screen "8_1" 800x480, template "Template_2"
   Button "Button_1" at 40,240 size 120x40; TextOff 'Acyclovir'
      on Click: ActivateScreen("4_ORDER", 0); SetTag("Selected_URL", 'file:///C:/ASRS_Video/clip291.html')
      on Activate: SetTag("Selected_Medicine", 291)
      on Release: SetTag("ยา 291", 0)
      on Press: SetTag("ยา 291", 1)
   Button "Button_10" at 40,416 size 120x40; TextOff 'Remdesivir'
      on Click: ActivateScreen("4_ORDER", 0); SetTag("Selected_URL", 'file:///C:/ASRS_Video/clip296.html')
      on Activate: SetTag("Selected_Medicine", 296)
      on Release: SetTag("ยา 296", 0)
      on Press: SetTag("ยา 296", 1)
   Button "Button_2" at 191,241 size 120x40; TextOff 'Valacyclovir'
      on Click: ActivateScreen("4_ORDER", 0); SetTag("Selected_URL", 'file:///C:/ASRS_Video/clip292.html')
      on Activate: SetTag("Selected_Medicine", 292)
      on Release: SetTag("ยา 292", 0)
      on Press: SetTag("ยา 292", 1)
   Button "Button_3" at 192,416 size 120x40; TextOff 'Favipiravir'
      on Click: ActivateScreen("4_ORDER", 0); SetTag("Selected_URL", 'file:///C:/ASRS_Video/clip297.html')
      on Activate: SetTag("Selected_Medicine", 297)
      on Release: SetTag("ยา 297", 0)
      on Press: SetTag("ยา 297", 1)
   Button "Button_4" at 342,241 size 120x40; TextOff 'Ganciclovir'
      on Click: ActivateScreen("4_ORDER", 0); SetTag("Selected_URL", 'file:///C:/ASRS_Video/clip293.html')
      on Activate: SetTag("Selected_Medicine", 293)
      on Release: SetTag("ยา 293", 0)
      on Press: SetTag("ยา 293", 1)
   Button "Button_5" at 342,417 size 120x40; TextOff 'Lamivudine'
      on Click: ActivateScreen("4_ORDER", 0); SetTag("Selected_URL", 'file:///C:/ASRS_Video/clip298.html')
      on Activate: SetTag("Selected_Medicine", 298)
      on Release: SetTag("ยา 298", 0)
      on Press: SetTag("ยา 298", 1)
   Button "Button_6" at 492,416 size 120x40; TextOff 'Zidovudine'
      on Click: ActivateScreen("4_ORDER", 0); SetTag("Selected_URL", 'file:///C:/ASRS_Video/clip299.html')
      on Activate: SetTag("Selected_Medicine", 299)
      on Release: SetTag("ยา 299", 0)
      on Press: SetTag("ยา 299", 1)
   Button "Button_7" at 492,240 size 120x40; TextOff 'Oseltamivir'
      on Click: ActivateScreen("4_ORDER", 0); SetTag("Selected_URL", 'file:///C:/ASRS_Video/clip294.html')
      on Activate: SetTag("Selected_Medicine", 294)
      on Release: SetTag("ยา 294", 0)
      on Press: SetTag("ยา 294", 1)
   Button "Button_8" at 644,240 size 120x40; TextOff 'Zanamivir'
      on Click: ActivateScreen("4_ORDER", 0); SetTag("Selected_URL", 'file:///C:/ASRS_Video/clip295.html')
      on Activate: SetTag("Selected_Medicine", 295)
      on Release: SetTag("ยา 295", 0)
      on Press: SetTag("ยา 295", 1)
   Button "Button_11" at 645,416 size 120x40; TextOff 'Tenofovir'
      on Click: ActivateScreen("4_ORDER", 0); SetTag("Selected_URL", 'file:///C:/ASRS_Video/clip300.html')
      on Activate: SetTag("Selected_Medicine", 300)
      on Release: SetTag("ยา 300", 0)
      on Press: SetTag("ยา 300", 1)
   Button "Button_12" at 24,16 size 94x40; TextOff 'Back'
      on Press: ActivateScreen("7_1", 0)
   Button "Button_9" at 688,16 size 96x40; TextOff 'Next'
      on Press: ActivateScreen("9_1", 0)
   GraphicView "Template_Graphic view_2" at 27,19 size 36x32; Picture "fast-backward"
   GraphicView "Template_Graphic view_1" at 693,20 size 36x32; Picture "play"
   GraphicView "Template_Graphic view_3" at 37,128 size 120x104; Picture "71"
   GraphicView "Template_Graphic view_4" at 191,129 size 120x104; Picture "72"
   GraphicView "Template_Graphic view_5" at 339,129 size 120x104; Picture "73"
   GraphicView "Template_Graphic view_6" at 493,129 size 120x104; Picture "74"
   GraphicView "Template_Graphic view_7" at 645,129 size 120x104; Picture "75"
   GraphicView "Template_Graphic view_8" at 38,305 size 120x104; Picture "76"
   GraphicView "Template_Graphic view_9" at 189,304 size 120x112; Picture "77"
   GraphicView "Template_Graphic view_10" at 351,307 size 96x104; Picture "78"
   GraphicView "Template_Graphic view_11" at 491,299 size 120x112; Picture "79"
   GraphicView "Template_Graphic view_12" at 645,304 size 120x104; Picture "80"
   TextField "Template_Text field_2" at 201,80 size 20x32; Text '8'

screen "9_1" 800x480, template "Template_2"
   Button "Button_1" at 38,239 size 120x40; TextOff 'Efavirenz'
      on Click: ActivateScreen("4_ORDER", 0); SetTag("Selected_URL", 'file:///C:/ASRS_Video/clip301.html')
      on Activate: SetTag("Selected_Medicine", 301)
      on Release: SetTag("ยา 301", 0)
      on Press: SetTag("ยา 301", 1)
   Button "Button_10" at 38,415 size 120x40; TextOff 'Mebendazole'
      on Click: ActivateScreen("4_ORDER", 0); SetTag("Selected_URL", 'file:///C:/ASRS_Video/clip306.html')
      on Activate: SetTag("Selected_Medicine", 306)
      on Release: SetTag("ยา 306", 0)
      on Press: SetTag("ยา 306", 1)
   Button "Button_2" at 189,240 size 120x40; TextOff 'Dolutegravir'
      on Click: ActivateScreen("4_ORDER", 0); SetTag("Selected_URL", 'file:///C:/ASRS_Video/clip302.html')
      on Activate: SetTag("Selected_Medicine", 302)
      on Release: SetTag("ยา 302", 0)
      on Press: SetTag("ยา 302", 1)
   Button "Button_3" at 190,415 size 120x40; TextOff 'Ivermectin'
      on Click: ActivateScreen("4_ORDER", 0); SetTag("Selected_URL", 'file:///C:/ASRS_Video/clip307.html')
      on Activate: SetTag("Selected_Medicine", 307)
      on Release: SetTag("ยา 307", 0)
      on Press: SetTag("ยา 307", 1)
   Button "Button_4" at 340,240 size 120x40; TextOff 'Nevirapine'
      on Click: ActivateScreen("4_ORDER", 0); SetTag("Selected_URL", 'file:///C:/ASRS_Video/clip303.html')
      on Activate: SetTag("Selected_Medicine", 303)
      on Release: SetTag("ยา 303", 0)
      on Press: SetTag("ยา 303", 1)
   Button "Button_5" at 340,416 size 120x40; TextOff 'Praziquantel'
      on Click: ActivateScreen("4_ORDER", 0); SetTag("Selected_URL", 'file:///C:/ASRS_Video/clip308.html')
      on Activate: SetTag("Selected_Medicine", 308)
      on Release: SetTag("ยา 308", 0)
      on Press: SetTag("ยา 308", 1)
   Button "Button_6" at 492,416 size 120x40; TextOff 'Pyrantel pamoate'
      on Click: ActivateScreen("4_ORDER", 0); SetTag("Selected_URL", 'file:///C:/ASRS_Video/clip309.html')
      on Activate: SetTag("Selected_Medicine", 309)
      on Release: SetTag("ยา 309", 0)
      on Press: SetTag("ยา 309", 1)
   Button "Button_7" at 492,240 size 120x40; TextOff 'Lopinavir ritonavir'
      on Click: ActivateScreen("4_ORDER", 0); SetTag("Selected_URL", 'file:///C:/ASRS_Video/clip304.html')
      on Activate: SetTag("Selected_Medicine", 304)
      on Release: SetTag("ยา 304", 0)
      on Press: SetTag("ยา 304", 1)
   Button "Button_8" at 644,240 size 120x40; TextOff 'Albendazole'
      on Click: ActivateScreen("4_ORDER", 0); SetTag("Selected_URL", 'file:///C:/ASRS_Video/clip305.html')
      on Activate: SetTag("Selected_Medicine", 305)
      on Release: SetTag("ยา 305", 0)
      on Press: SetTag("ยา 305", 1)
   Button "Button_11" at 645,416 size 120x40; TextOff 'Diethylcarbamazine'
      on Click: ActivateScreen("4_ORDER", 0); SetTag("Selected_URL", 'file:///C:/ASRS_Video/clip310.html')
      on Activate: SetTag("Selected_Medicine", 310)
      on Release: SetTag("ยา 310", 0)
      on Press: SetTag("ยา 310", 1)
   Button "Button_12" at 24,16 size 94x40; TextOff 'Back'
      on Press: ActivateScreen("8_1", 0)
   Button "Button_9" at 688,16 size 96x40; TextOff 'Next'
      on Press: ActivateScreen("10_1", 0)
   GraphicView "Template_Graphic view_2" at 27,19 size 36x32; Picture "fast-backward"
   GraphicView "Template_Graphic view_1" at 693,20 size 36x32; Picture "play"
   GraphicView "Template_Graphic view_3" at 37,128 size 120x104; Picture "81"
   GraphicView "Template_Graphic view_4" at 191,129 size 120x104; Picture "82"
   GraphicView "Template_Graphic view_5" at 339,129 size 120x104; Picture "83"
   GraphicView "Template_Graphic view_6" at 493,129 size 120x104; Picture "84"
   GraphicView "Template_Graphic view_7" at 645,129 size 120x104; Picture "85"
   GraphicView "Template_Graphic view_8" at 38,305 size 120x104; Picture "86"
   GraphicView "Template_Graphic view_9" at 189,304 size 120x112; Picture "87"
   GraphicView "Template_Graphic view_10" at 351,307 size 96x104; Picture "88"
   GraphicView "Template_Graphic view_11" at 497,304 size 120x112; Picture "89"
   GraphicView "Template_Graphic view_12" at 645,304 size 120x104; Picture "90"
   TextField "Template_Text field_2" at 201,80 size 20x32; Text '9'

screen "10_1" 800x480, template "Template_2"
   Button "Button_1" at 38,239 size 120x40; TextOff 'Chloroquine'
      on Click: ActivateScreen("4_ORDER", 0); SetTag("Selected_URL", 'file:///C:/ASRS_Video/clip311.html')
      on Activate: SetTag("Selected_Medicine", 311)
      on Release: SetTag("ยา 311", 0)
      on Press: SetTag("ยา 311", 1)
   Button "Button_10" at 38,415 size 120x40; TextOff 'Dapsone'
      on Click: ActivateScreen("4_ORDER", 0); SetTag("Selected_URL", 'file:///C:/ASRS_Video/clip316.html')
      on Activate: SetTag("Selected_Medicine", 316)
      on Release: SetTag("ยา 316", 0)
      on Press: SetTag("ยา 316", 1)
   Button "Button_2" at 189,240 size 120x40; TextOff 'Primaquine'
      on Click: ActivateScreen("4_ORDER", 0); SetTag("Selected_URL", 'file:///C:/ASRS_Video/clip312.html')
      on Activate: SetTag("Selected_Medicine", 312)
      on Release: SetTag("ยา 312", 0)
      on Press: SetTag("ยา 312", 1)
   Button "Button_3" at 190,415 size 120x40; TextOff 'Permethrin'
      on Click: ActivateScreen("4_ORDER", 0); SetTag("Selected_URL", 'file:///C:/ASRS_Video/clip317.html')
      on Activate: SetTag("Selected_Medicine", 317)
      on Release: SetTag("ยา 317", 0)
      on Press: SetTag("ยา 317", 1)
   Button "Button_4" at 340,240 size 120x40; TextOff 'Artesunate'
      on Click: ActivateScreen("4_ORDER", 0); SetTag("Selected_URL", 'file:///C:/ASRS_Video/clip313.html')
      on Activate: SetTag("Selected_Medicine", 313)
      on Release: SetTag("ยา 313", 0)
      on Press: SetTag("ยา 313", 1)
   Button "Button_5" at 340,416 size 120x40; TextOff 'Benzyl benzoate'
      on Click: ActivateScreen("4_ORDER", 0); SetTag("Selected_URL", 'file:///C:/ASRS_Video/clip318.html')
      on Activate: SetTag("Selected_Medicine", 318)
      on Release: SetTag("ยา 318", 0)
      on Press: SetTag("ยา 318", 1)
   Button "Button_6" at 492,416 size 120x40; TextOff 'Povidone iodine'
      on Click: ActivateScreen("4_ORDER", 0); SetTag("Selected_URL", 'file:///C:/ASRS_Video/clip319.html')
      on Activate: SetTag("Selected_Medicine", 319)
      on Release: SetTag("ยา 319", 0)
      on Press: SetTag("ยา 319", 1)
   Button "Button_7" at 492,240 size 120x40; TextOff 'Artemether lumefantrine'
      on Click: ActivateScreen("4_ORDER", 0); SetTag("Selected_URL", 'file:///C:/ASRS_Video/clip314.html')
      on Activate: SetTag("Selected_Medicine", 314)
      on Release: SetTag("ยา 314", 0)
      on Press: SetTag("ยา 314", 1)
   Button "Button_8" at 644,240 size 120x40; TextOff 'Quinine'
      on Click: ActivateScreen("4_ORDER", 0); SetTag("Selected_URL", 'file:///C:/ASRS_Video/clip315.html')
      on Activate: SetTag("Selected_Medicine", 315)
      on Release: SetTag("ยา 315", 0)
      on Press: SetTag("ยา 315", 1)
   Button "Button_11" at 645,416 size 120x40; TextOff 'Chlorhexidine'
      on Click: ActivateScreen("4_ORDER", 0); SetTag("Selected_URL", 'file:///C:/ASRS_Video/clip320.html')
      on Activate: SetTag("Selected_Medicine", 320)
      on Release: SetTag("ยา 320", 0)
      on Press: SetTag("ยา 320", 1)
   Button "Button_12" at 24,16 size 94x40; TextOff 'Back'
      on Press: ActivateScreen("9_1", 0)
   Button "Button_9" at 688,16 size 96x40; TextOff 'Next'
      on Press: ActivateScreen("11_1", 0)
   GraphicView "Template_Graphic view_2" at 27,19 size 36x32; Picture "fast-backward"
   GraphicView "Template_Graphic view_1" at 693,20 size 36x32; Picture "play"
   GraphicView "Template_Graphic view_3" at 37,128 size 120x104; Picture "91"
   GraphicView "Template_Graphic view_4" at 191,129 size 120x104; Picture "92"
   GraphicView "Template_Graphic view_5" at 339,129 size 120x104; Picture "93"
   GraphicView "Template_Graphic view_6" at 493,129 size 120x104; Picture "94"
   GraphicView "Template_Graphic view_7" at 645,129 size 120x104; Picture "95"
   GraphicView "Template_Graphic view_8" at 38,305 size 120x104; Picture "96"
   GraphicView "Template_Graphic view_9" at 189,304 size 120x112; Picture "97"
   GraphicView "Template_Graphic view_10" at 351,307 size 96x104; Picture "98"
   GraphicView "Template_Graphic view_11" at 497,304 size 104x104; Picture "99"
   GraphicView "Template_Graphic view_12" at 645,304 size 120x104; Picture "100"
   TextField "Template_Text field_2" at 201,80 size 36x32; Text '10'

screen "11_1" 800x480, template "Template_2"
   Button "Button_1" at 38,239 size 120x40; TextOff 'Colistin'
      on Click: ActivateScreen("4_ORDER", 0); SetTag("Selected_URL", 'file:///C:/ASRS_Video/clip321.html')
      on Activate: SetTag("Selected_Medicine", 321)
      on Release: SetTag("ยา 321", 0)
      on Press: SetTag("ยา 321", 1)
   Button "Button_10" at 38,415 size 120x40; TextOff 'Rabies vaccine'
      on Click: ActivateScreen("4_ORDER", 0); SetTag("Selected_URL", 'file:///C:/ASRS_Video/clip326.html')
      on Activate: SetTag("Selected_Medicine", 326)
      on Release: SetTag("ยา 326", 0)
      on Press: SetTag("ยา 326", 1)
   Button "Button_2" at 189,240 size 120x40; TextOff 'Caspofungin'
      on Click: ActivateScreen("4_ORDER", 0); SetTag("Selected_URL", 'file:///C:/ASRS_Video/clip322.html')
      on Activate: SetTag("Selected_Medicine", 322)
      on Release: SetTag("ยา 322", 0)
      on Press: SetTag("ยา 322", 1)
   Button "Button_3" at 190,415 size 120x40; TextOff 'Influenza vaccine'
      on Click: ActivateScreen("4_ORDER", 0); SetTag("Selected_URL", 'file:///C:/ASRS_Video/clip327.html')
      on Activate: SetTag("Selected_Medicine", 327)
      on Release: SetTag("ยา 327", 0)
      on Press: SetTag("ยา 327", 1)
   Button "Button_4" at 340,240 size 120x40; TextOff 'Bacitracin'
      on Click: ActivateScreen("4_ORDER", 0); SetTag("Selected_URL", 'file:///C:/ASRS_Video/clip323.html')
      on Activate: SetTag("Selected_Medicine", 323)
      on Release: SetTag("ยา 323", 0)
      on Press: SetTag("ยา 323", 1)
   Button "Button_5" at 340,416 size 120x40; TextOff 'Hepatitis B vaccine'
      on Click: ActivateScreen("4_ORDER", 0); SetTag("Selected_URL", 'file:///C:/ASRS_Video/clip328.html')
      on Activate: SetTag("Selected_Medicine", 328)
      on Release: SetTag("ยา 328", 0)
      on Press: SetTag("ยา 328", 1)
   Button "Button_6" at 492,416 size 120x40; TextOff 'BCG vaccine'
      on Click: ActivateScreen("4_ORDER", 0); SetTag("Selected_URL", 'file:///C:/ASRS_Video/clip329.html')
      on Activate: SetTag("Selected_Medicine", 329)
      on Release: SetTag("ยา 329", 0)
      on Press: SetTag("ยา 329", 1)
   Button "Button_7" at 492,240 size 120x40; TextOff 'Fusidic acid'
      on Click: ActivateScreen("4_ORDER", 0); SetTag("Selected_URL", 'file:///C:/ASRS_Video/clip324.html')
      on Activate: SetTag("Selected_Medicine", 324)
      on Release: SetTag("ยา 324", 0)
      on Press: SetTag("ยา 324", 1)
   Button "Button_8" at 644,240 size 120x40; TextOff 'Mupirocin'
      on Click: ActivateScreen("4_ORDER", 0); SetTag("Selected_URL", 'file:///C:/ASRS_Video/clip325.html')
      on Activate: SetTag("Selected_Medicine", 325)
      on Release: SetTag("ยา 325", 0)
      on Press: SetTag("ยา 325", 1)
   Button "Button_11" at 645,416 size 120x40; TextOff 'DTP vaccine'
      on Click: ActivateScreen("4_ORDER", 0); SetTag("Selected_URL", 'file:///C:/ASRS_Video/clip330.html')
      on Activate: SetTag("Selected_Medicine", 330)
      on Release: SetTag("ยา 330", 0)
      on Press: SetTag("ยา 330", 1)
   Button "Button_12" at 24,16 size 94x40; TextOff 'Back'
      on Press: ActivateScreen("10_1", 0)
   Button "Button_9" at 688,16 size 96x40; TextOff 'Next'
      on Press: ActivateScreen("12_1", 0)
   GraphicView "Template_Graphic view_2" at 27,19 size 36x32; Picture "fast-backward"
   GraphicView "Template_Graphic view_1" at 693,20 size 36x32; Picture "play"
   GraphicView "Template_Graphic view_3" at 37,128 size 120x104; Picture "101"
   GraphicView "Template_Graphic view_4" at 191,129 size 120x104; Picture "102"
   GraphicView "Template_Graphic view_5" at 339,129 size 120x104; Picture "103"
   GraphicView "Template_Graphic view_6" at 493,129 size 120x104; Picture "104"
   GraphicView "Template_Graphic view_7" at 645,129 size 120x104; Picture "105"
   GraphicView "Template_Graphic view_8" at 38,305 size 120x104; Picture "106"
   GraphicView "Template_Graphic view_9" at 189,304 size 120x104; Picture "107"
   GraphicView "Template_Graphic view_10" at 351,307 size 96x104; Picture "108"
   GraphicView "Template_Graphic view_11" at 497,304 size 112x104; Picture "109"
   GraphicView "Template_Graphic view_12" at 645,304 size 120x104; Picture "110"
   TextField "Template_Text field_2" at 201,80 size 36x32; Text '11'

screen "12_1" 800x480, template "Template_2"
   Button "Button_1" at 38,239 size 120x40; TextOff 'MMR vaccine'
      on Click: ActivateScreen("4_ORDER", 0); SetTag("Selected_URL", 'file:///C:/ASRS_Video/clip331.html')
      on Activate: SetTag("Selected_Medicine", 331)
      on Release: SetTag("ยา 331", 0)
      on Press: SetTag("ยา 331", 1)
   Button "Button_10" at 38,415 size 120x40; TextOff 'Rotavirus vaccine'
      on Click: ActivateScreen("4_ORDER", 0); SetTag("Selected_URL", 'file:///C:/ASRS_Video/clip336.html')
      on Activate: SetTag("Selected_Medicine", 336)
      on Release: SetTag("ยา 336", 0)
      on Press: SetTag("ยา 336", 1)
   Button "Button_2" at 189,240 size 120x40; TextOff 'JE vaccine'
      on Click: ActivateScreen("4_ORDER", 0); SetTag("Selected_URL", 'file:///C:/ASRS_Video/clip332.html')
      on Activate: SetTag("Selected_Medicine", 332)
      on Release: SetTag("ยา 332", 0)
      on Press: SetTag("ยา 332", 1)
   Button "Button_3" at 190,415 size 120x40; TextOff 'COVID-19 vaccine'
      on Click: ActivateScreen("4_ORDER", 0); SetTag("Selected_URL", 'file:///C:/ASRS_Video/clip337.html')
      on Activate: SetTag("Selected_Medicine", 337)
      on Release: SetTag("ยา 337", 0)
      on Press: SetTag("ยา 337", 1)
   Button "Button_4" at 340,240 size 120x40; TextOff 'HPV vaccine'
      on Click: ActivateScreen("4_ORDER", 0); SetTag("Selected_URL", 'file:///C:/ASRS_Video/clip333.html')
      on Activate: SetTag("Selected_Medicine", 333)
      on Release: SetTag("ยา 333", 0)
      on Press: SetTag("ยา 333", 1)
   Button "Button_5" at 340,416 size 120x40; TextOff 'Tetanus toxoid'
      on Click: ActivateScreen("4_ORDER", 0); SetTag("Selected_URL", 'file:///C:/ASRS_Video/clip338.html')
      on Activate: SetTag("Selected_Medicine", 338)
      on Release: SetTag("ยา 338", 0)
      on Press: SetTag("ยา 338", 1)
   Button "Button_6" at 492,416 size 120x40; TextOff 'Rabies immunoglobulin'
      on Click: ActivateScreen("4_ORDER", 0); SetTag("Selected_URL", 'file:///C:/ASRS_Video/clip339.html')
      on Activate: SetTag("Selected_Medicine", 339)
      on Release: SetTag("ยา 339", 0)
      on Press: SetTag("ยา 339", 1)
   Button "Button_7" at 492,240 size 120x40; TextOff 'Varicella vaccine'
      on Click: ActivateScreen("4_ORDER", 0); SetTag("Selected_URL", 'file:///C:/ASRS_Video/clip334.html')
      on Activate: SetTag("Selected_Medicine", 334)
      on Release: SetTag("ยา 334", 0)
      on Press: SetTag("ยา 334", 1)
   Button "Button_8" at 644,240 size 120x40; TextOff 'Pneumococcal vaccine'
      on Click: ActivateScreen("4_ORDER", 0); SetTag("Selected_URL", 'file:///C:/ASRS_Video/clip335.html')
      on Activate: SetTag("Selected_Medicine", 335)
      on Release: SetTag("ยา 335", 0)
      on Press: SetTag("ยา 335", 1)
   Button "Button_11" at 645,416 size 120x40; TextOff 'Hepatitis B immunoglobulin'
      on Click: ActivateScreen("4_ORDER", 0); SetTag("Selected_URL", 'file:///C:/ASRS_Video/clip340.html')
      on Activate: SetTag("Selected_Medicine", 340)
      on Release: SetTag("ยา 340", 0)
      on Press: SetTag("ยา 340", 1)
   Button "Button_12" at 24,16 size 94x40; TextOff 'Back'
      on Press: ActivateScreen("11_1", 0)
   GraphicView "Template_Graphic view_2" at 27,19 size 36x32; Picture "fast-backward"
   GraphicView "Template_Graphic view_3" at 37,128 size 120x104; Picture "111"
   GraphicView "Template_Graphic view_4" at 191,129 size 120x104; Picture "112"
   GraphicView "Template_Graphic view_5" at 339,129 size 120x104; Picture "113"
   GraphicView "Template_Graphic view_6" at 493,129 size 120x104; Picture "114"
   GraphicView "Template_Graphic view_7" at 645,129 size 120x104; Picture "115"
   GraphicView "Template_Graphic view_8" at 38,305 size 120x104; Picture "116"
   GraphicView "Template_Graphic view_9" at 189,304 size 120x112; Picture "117"
   GraphicView "Template_Graphic view_10" at 351,307 size 96x104; Picture "118"
   GraphicView "Template_Graphic view_11" at 497,304 size 120x112; Picture "119"
   GraphicView "Template_Graphic view_12" at 645,304 size 120x104; Picture "120"
   TextField "Template_Text field_2" at 201,80 size 36x32; Text '12'

screen "1-10" 800x480, template "Template_2"
   Button "Button_1" at 40,240 size 120x40; TextOff 'Lidocaine'
      on Click: ActivateScreen("4_ORDER", 0); SetTag("Selected_URL", 'file:///C:/ASRS_Video/clip1.html')
      on Activate: SetTag("Selected_Medicine", 1)
      on Release: SetTag("ยา 1", 0)
      on Press: SetTag("ยา 1", 1)
   Button "Button_10" at 38,415 size 120x40; TextOff 'Tetracaine'
      on Click: ActivateScreen("4_ORDER", 0); SetTag("Selected_URL", 'file:///C:/ASRS_Video/clip6.html')
      on Activate: SetTag("Selected_Medicine", 6)
      on Release: SetTag("ยา 6", 0)
      on Press: SetTag("ยา 6", 1)
   Button "Button_2" at 189,240 size 120x40; TextOff 'Bupivacaine'
      on Click: ActivateScreen("4_ORDER", 0); SetTag("Selected_URL", 'file:///C:/ASRS_Video/clip2.html')
      on Activate: SetTag("Selected_Medicine", 2)
      on Release: SetTag("ยา 2", 0)
      on Press: SetTag("ยา 2", 1)
   Button "Button_3" at 190,415 size 120x40; TextOff 'Propofol'
      on Click: ActivateScreen("4_ORDER", 0); SetTag("Selected_URL", 'file:///C:/ASRS_Video/clip7.html')
      on Activate: SetTag("Selected_Medicine", 7)
      on Release: SetTag("ยา 7", 0)
      on Press: SetTag("ยา 7", 1)
   Button "Button_4" at 340,240 size 120x40; TextOff 'Ropivacaine'
      on Click: ActivateScreen("4_ORDER", 0); SetTag("Selected_URL", 'file:///C:/ASRS_Video/clip3.html')
      on Activate: SetTag("Selected_Medicine", 3)
      on Release: SetTag("ยา 3", 0)
      on Press: SetTag("ยา 3", 1)
   Button "Button_5" at 340,416 size 120x40; TextOff 'Ketamine'
      on Click: ActivateScreen("4_ORDER", 0); SetTag("Selected_URL", 'file:///C:/ASRS_Video/clip8.html')
      on Activate: SetTag("Selected_Medicine", 8)
      on Release: SetTag("ยา 8", 0)
      on Press: SetTag("ยา 8", 1)
   Button "Button_6" at 492,416 size 120x40; TextOff 'Etomidate'
      on Click: ActivateScreen("4_ORDER", 0); SetTag("Selected_URL", 'file:///C:/ASRS_Video/clip9.html')
      on Activate: SetTag("Selected_Medicine", 9)
      on Release: SetTag("ยา 9", 0)
      on Press: SetTag("ยา 9", 1)
   Button "Button_7" at 492,240 size 120x40; TextOff 'Procaine'
      on Click: ActivateScreen("4_ORDER", 0); SetTag("Selected_URL", 'file:///C:/ASRS_Video/clip4.html')
      on Activate: SetTag("Selected_Medicine", 4)
      on Release: SetTag("ยา 4", 0)
      on Press: SetTag("ยา 4", 1)
   Button "Button_8" at 644,240 size 120x40; TextOff 'Benzocaine'
      on Click: ActivateScreen("4_ORDER", 0); SetTag("Selected_URL", 'file:///C:/ASRS_Video/clip5.html')
      on Activate: SetTag("Selected_Medicine", 5)
      on Release: SetTag("ยา 5", 0)
      on Press: SetTag("ยา 5", 1)
   Button "Button_11" at 645,416 size 120x40; TextOff 'Thiopental'
      on Click: ActivateScreen("4_ORDER", 0); SetTag("Selected_URL", 'file:///C:/ASRS_Video/clip10.html')
      on Activate: SetTag("Selected_Medicine", 10)
      on Release: SetTag("ยา 10", 0)
      on Press: SetTag("ยา 10", 1)
   Button "Button_12" at 688,16 size 96x40; TextOff 'Next'
      on Press: ActivateScreen("11-20", 0)
   Button "Button_9" at 24,16 size 94x40; TextOff 'Back'
      on Press: ActivateScreen("4_ORDER", 0)
   GraphicView "Template_Graphic view_2" at 693,20 size 36x32; Picture "play"
   GraphicView "Template_Graphic view_1" at 27,19 size 36x32; Picture "fast-backward"
   GraphicView "Template_Graphic view_3" at 38,127 size 120x112; Picture "Picture1"
   GraphicView "Template_Graphic view_4" at 190,128 size 120x112; Picture "Picture2"
   GraphicView "Template_Graphic view_5" at 340,128 size 120x112; Picture "Picture3"
   GraphicView "Template_Graphic view_6" at 493,128 size 120x112; Picture "Picture4"
   GraphicView "Template_Graphic view_7" at 644,128 size 120x112; Picture "Picture5"
   GraphicView "Template_Graphic view_8" at 37,302 size 120x112; Picture "Picture6"
   GraphicView "Template_Graphic view_9" at 189,303 size 120x112; Picture "Picture7"
   GraphicView "Template_Graphic view_10" at 339,303 size 120x112; Picture "Picture8"
   GraphicView "Template_Graphic view_11" at 492,303 size 120x112; Picture "Picture9"
   GraphicView "Template_Graphic view_12" at 643,303 size 120x112; Picture "Picture10"
   TextField "Template_Text field_2" at 201,80 size 20x32; Text '1'

screen "11-20" 800x480, template "Template_2"
   Button "Button_1" at 38,239 size 120x40; TextOff 'Midazolam'
      on Click: ActivateScreen("4_ORDER", 0); SetTag("Selected_URL", 'file:///C:/ASRS_Video/clip11.html')
      on Activate: SetTag("Selected_Medicine", 11)
      on Release: SetTag("ยา 11", 0)
      on Press: SetTag("ยา 11", 1)
   Button "Button_9" at 688,16 size 96x40; TextOff 'Next'
      on Press: ActivateScreen("21-30", 0)
   Button "Button_10" at 38,415 size 120x40; TextOff 'Pethidine'
      on Click: ActivateScreen("4_ORDER", 0); SetTag("Selected_URL", 'file:///C:/ASRS_Video/clip16.html')
      on Activate: SetTag("Selected_Medicine", 16)
      on Release: SetTag("ยา 16", 0)
      on Press: SetTag("ยา 16", 1)
   Button "Button_2" at 189,240 size 120x40; TextOff 'Diazepam'
      on Click: ActivateScreen("4_ORDER", 0); SetTag("Selected_URL", 'file:///C:/ASRS_Video/clip12.html')
      on Activate: SetTag("Selected_Medicine", 12)
      on Release: SetTag("ยา 12", 0)
      on Press: SetTag("ยา 12", 1)
   Button "Button_3" at 190,415 size 120x40; TextOff 'Tramadol'
      on Click: ActivateScreen("4_ORDER", 0); SetTag("Selected_URL", 'file:///C:/ASRS_Video/clip17.html')
      on Activate: SetTag("Selected_Medicine", 17)
      on Release: SetTag("ยา 17", 0)
      on Press: SetTag("ยา 17", 1)
   Button "Button_4" at 340,240 size 120x40; TextOff 'Lorazepam'
      on Click: ActivateScreen("4_ORDER", 0); SetTag("Selected_URL", 'file:///C:/ASRS_Video/clip13.html')
      on Activate: SetTag("Selected_Medicine", 13)
      on Release: SetTag("ยา 13", 0)
      on Press: SetTag("ยา 13", 1)
   Button "Button_5" at 340,416 size 120x40; TextOff 'Nalbuphine'
      on Click: ActivateScreen("4_ORDER", 0); SetTag("Selected_URL", 'file:///C:/ASRS_Video/clip18.html')
      on Activate: SetTag("Selected_Medicine", 18)
      on Release: SetTag("ยา 18", 0)
      on Press: SetTag("ยา 18", 1)
   Button "Button_6" at 492,416 size 120x40; TextOff 'Remifentanil'
      on Click: ActivateScreen("4_ORDER", 0); SetTag("Selected_URL", 'file:///C:/ASRS_Video/clip19.html')
      on Activate: SetTag("Selected_Medicine", 19)
      on Release: SetTag("ยา 19", 0)
      on Press: SetTag("ยา 19", 1)
   Button "Button_7" at 492,240 size 120x40; TextOff 'Fentanyl'
      on Click: ActivateScreen("4_ORDER", 0); SetTag("Selected_URL", 'file:///C:/ASRS_Video/clip14.html')
      on Activate: SetTag("Selected_Medicine", 14)
      on Release: SetTag("ยา 14", 0)
      on Press: SetTag("ยา 14", 1)
   Button "Button_8" at 644,240 size 120x40; TextOff 'Morphine'
      on Click: ActivateScreen("4_ORDER", 0); SetTag("Selected_URL", 'file:///C:/ASRS_Video/clip15.html')
      on Activate: SetTag("Selected_Medicine", 15)
      on Release: SetTag("ยา 15", 0)
      on Press: SetTag("ยา 15", 1)
   Button "Button_11" at 645,416 size 120x40; TextOff 'Succinylcholine'
      on Click: ActivateScreen("4_ORDER", 0); SetTag("Selected_URL", 'file:///C:/ASRS_Video/clip20.html')
      on Activate: SetTag("Selected_Medicine", 20)
      on Release: SetTag("ยา 20", 0)
      on Press: SetTag("ยา 20", 1)
   Button "Button_12" at 24,16 size 94x40; TextOff 'Back'
      on Press: ActivateScreen("1-10", 0)
   GraphicView "Template_Graphic view_1" at 693,20 size 36x32; Picture "play"
   GraphicView "Template_Graphic view_2" at 27,19 size 36x32; Picture "fast-backward"
   GraphicView "Template_Graphic view_3" at 38,127 size 120x112; Picture "Picture11"
   GraphicView "Template_Graphic view_4" at 190,128 size 120x104; Picture "Picture12"
   GraphicView "Template_Graphic view_5" at 340,128 size 120x104; Picture "Picture13"
   GraphicView "Template_Graphic view_6" at 493,128 size 120x112; Picture "Picture14"
   GraphicView "Template_Graphic view_7" at 644,128 size 120x112; Picture "Picture15"
   GraphicView "Template_Graphic view_8" at 37,302 size 120x112; Picture "Picture16"
   GraphicView "Template_Graphic view_9" at 189,303 size 120x112; Picture "Picture17"
   GraphicView "Template_Graphic view_10" at 339,303 size 120x112; Picture "Picture18"
   GraphicView "Template_Graphic view_11" at 492,303 size 120x112; Picture "Picture19"
   GraphicView "Template_Graphic view_12" at 643,303 size 120x112; Picture "Picture20"
   TextField "Template_Text field_2" at 201,80 size 20x32; Text '2'

screen "21-30" 800x480, template "Template_2"
   Button "Button_1" at 38,239 size 120x40; TextOff 'Rocuronium'
      on Click: ActivateScreen("4_ORDER", 0); SetTag("Selected_URL", 'file:///C:/ASRS_Video/clip21.html')
      on Activate: SetTag("Selected_Medicine", 21)
      on Release: SetTag("ยา 21", 0)
      on Press: SetTag("ยา 21", 1)
   Button "Button_9" at 688,16 size 96x40; TextOff 'Next'
      on Press: ActivateScreen("31-40", 0)
   Button "Button_10" at 38,415 size 120x40; TextOff 'Atropine'
      on Click: ActivateScreen("4_ORDER", 0); SetTag("Selected_URL", 'file:///C:/ASRS_Video/clip26.html')
      on Activate: SetTag("Selected_Medicine", 26)
      on Release: SetTag("ยา 26", 0)
      on Press: SetTag("ยา 26", 1)
   Button "Button_2" at 189,240 size 120x40; TextOff 'Vecuronium'
      on Click: ActivateScreen("4_ORDER", 0); SetTag("Selected_URL", 'file:///C:/ASRS_Video/clip22.html')
      on Activate: SetTag("Selected_Medicine", 22)
      on Release: SetTag("ยา 21", 0)
      on Press: SetTag("ยา 22", 1)
   Button "Button_3" at 190,415 size 120x40; TextOff 'Glycopyrrolate'
      on Click: ActivateScreen("4_ORDER", 0); SetTag("Selected_URL", 'file:///C:/ASRS_Video/clip27.html')
      on Activate: SetTag("Selected_Medicine", 27)
      on Release: SetTag("ยา 27", 0)
      on Press: SetTag("ยา 27", 1)
   Button "Button_4" at 340,240 size 120x40; TextOff 'Atracurium'
      on Click: ActivateScreen("4_ORDER", 0); SetTag("Selected_URL", 'file:///C:/ASRS_Video/clip23.html')
      on Activate: SetTag("Selected_Medicine", 23)
      on Release: SetTag("ยา 23", 0)
      on Press: SetTag("ยา 23", 1)
   Button "Button_5" at 340,416 size 120x40; TextOff 'Epinephrine'
      on Click: ActivateScreen("4_ORDER", 0); SetTag("Selected_URL", 'file:///C:/ASRS_Video/clip28.html')
      on Activate: SetTag("Selected_Medicine", 28)
      on Release: SetTag("ยา 28", 0)
      on Press: SetTag("ยา 28", 1)
   Button "Button_6" at 492,416 size 120x40; TextOff 'Norepinephrine'
      on Click: ActivateScreen("4_ORDER", 0); SetTag("Selected_URL", 'file:///C:/ASRS_Video/clip29.html')
      on Activate: SetTag("Selected_Medicine", 29)
      on Release: SetTag("ยา 29", 0)
      on Press: SetTag("ยา 29", 1)
   Button "Button_7" at 492,240 size 120x40; TextOff 'Cisatracurium'
      on Click: ActivateScreen("4_ORDER", 0); SetTag("Selected_URL", 'file:///C:/ASRS_Video/clip24.html')
      on Activate: SetTag("Selected_Medicine", 24)
      on Release: SetTag("ยา 24", 0)
      on Press: SetTag("ยา 24", 1)
   Button "Button_8" at 644,240 size 120x40; TextOff 'Neostigmine'
      on Click: ActivateScreen("4_ORDER", 0); SetTag("Selected_URL", 'file:///C:/ASRS_Video/clip25.html')
      on Activate: SetTag("Selected_Medicine", 25)
      on Release: SetTag("ยา 25", 0)
      on Press: SetTag("ยา 25", 1)
   Button "Button_11" at 645,416 size 120x40; TextOff 'Dopamine'
      on Click: ActivateScreen("4_ORDER", 0); SetTag("Selected_URL", 'file:///C:/ASRS_Video/clip30.html')
      on Activate: SetTag("Selected_Medicine", 30)
      on Release: SetTag("ยา 30", 0)
      on Press: SetTag("ยา 30", 1)
   Button "Button_12" at 24,16 size 94x40; TextOff 'Back'
      on Press: ActivateScreen("11-20", 0)
   GraphicView "Template_Graphic view_1" at 693,20 size 36x32; Picture "play"
   GraphicView "Template_Graphic view_2" at 27,19 size 36x32; Picture "fast-backward"
   GraphicView "Template_Graphic view_3" at 38,127 size 120x112; Picture "Picture21"
   GraphicView "Template_Graphic view_4" at 190,128 size 120x112; Picture "Picture22"
   GraphicView "Template_Graphic view_5" at 340,128 size 120x112; Picture "Picture23"
   GraphicView "Template_Graphic view_6" at 493,128 size 120x112; Picture "Picture24"
   GraphicView "Template_Graphic view_7" at 644,128 size 120x112; Picture "Picture25"
   GraphicView "Template_Graphic view_8" at 37,302 size 120x112; Picture "Picture26"
   GraphicView "Template_Graphic view_9" at 189,303 size 120x112; Picture "Picture27"
   GraphicView "Template_Graphic view_10" at 339,303 size 120x112; Picture "Picture28"
   GraphicView "Template_Graphic view_11" at 492,303 size 120x112; Picture "Picture29"
   GraphicView "Template_Graphic view_12" at 643,303 size 120x112; Picture "Picture30"
   TextField "Template_Text field_2" at 201,80 size 20x32; Text '3'

screen "31-40" 800x480, template "Template_2"
   Button "Button_1" at 38,239 size 120x40; TextOff 'Dobutamine'
      on Click: ActivateScreen("4_ORDER", 0); SetTag("Selected_URL", 'file:///C:/ASRS_Video/clip31.html')
      on Activate: SetTag("Selected_Medicine", 31)
      on Release: SetTag("ยา 31", 0)
      on Press: SetTag("ยา 31", 1)
   Button "Button_9" at 688,16 size 96x40; TextOff 'Next'
      on Press: ActivateScreen("41-50", 0)
   Button "Button_10" at 38,415 size 120x40; TextOff 'Amiodarone'
      on Click: ActivateScreen("4_ORDER", 0); SetTag("Selected_URL", 'file:///C:/ASRS_Video/clip36.html')
      on Activate: SetTag("Selected_Medicine", 36)
      on Release: SetTag("ยา 36", 0)
      on Press: SetTag("ยา 36", 1)
   Button "Button_2" at 189,240 size 120x40; TextOff 'Phenylephrine'
      on Click: ActivateScreen("4_ORDER", 0); SetTag("Selected_URL", 'file:///C:/ASRS_Video/clip32.html')
      on Activate: SetTag("Selected_Medicine", 32)
      on Release: SetTag("ยา 32", 0)
      on Press: SetTag("ยา 32", 1)
   Button "Button_3" at 190,415 size 120x40; TextOff 'Adenosine'
      on Click: ActivateScreen("4_ORDER", 0); SetTag("Selected_URL", 'file:///C:/ASRS_Video/clip37.html')
      on Activate: SetTag("Selected_Medicine", 37)
      on Release: SetTag("ยา 37", 0)
      on Press: SetTag("ยา 37", 1)
   Button "Button_4" at 340,240 size 120x40; TextOff 'Vasopressin'
      on Click: ActivateScreen("4_ORDER", 0); SetTag("Selected_URL", 'file:///C:/ASRS_Video/clip33.html')
      on Activate: SetTag("Selected_Medicine", 33)
      on Release: SetTag("ยา 33", 0)
      on Press: SetTag("ยา 33", 1)
   Button "Button_5" at 340,416 size 120x40; TextOff 'Verapamil'
      on Click: ActivateScreen("4_ORDER", 0); SetTag("Selected_URL", 'file:///C:/ASRS_Video/clip38.html')
      on Activate: SetTag("Selected_Medicine", 38)
      on Release: SetTag("ยา 38", 0)
      on Press: SetTag("ยา 38", 1)
   Button "Button_6" at 492,416 size 120x40; TextOff 'Diltiazem'
      on Click: ActivateScreen("4_ORDER", 0); SetTag("Selected_URL", 'file:///C:/ASRS_Video/clip39.html')
      on Activate: SetTag("Selected_Medicine", 39)
      on Release: SetTag("ยา 39", 0)
      on Press: SetTag("ยา 39", 1)
   Button "Button_7" at 492,240 size 120x40; TextOff 'Nitroglycerin'
      on Click: ActivateScreen("4_ORDER", 0); SetTag("Selected_URL", 'file:///C:/ASRS_Video/clip34.html')
      on Activate: SetTag("Selected_Medicine", 34)
      on Release: SetTag("ยา 34", 0)
      on Press: SetTag("ยา 34", 1)
   Button "Button_8" at 644,240 size 120x40; TextOff 'Sodium nitroprusside'
      on Click: ActivateScreen("4_ORDER", 0); SetTag("Selected_URL", 'file:///C:/ASRS_Video/clip35.html')
      on Activate: SetTag("Selected_Medicine", 35)
      on Release: SetTag("ยา 35", 0)
      on Press: SetTag("ยา 35", 1)
   Button "Button_11" at 645,416 size 120x40; TextOff 'Lidocaine'
      on Click: ActivateScreen("4_ORDER", 0); SetTag("Selected_URL", 'file:///C:/ASRS_Video/clip40.html')
      on Activate: SetTag("Selected_Medicine", 40)
      on Release: SetTag("ยา 40", 0)
      on Press: SetTag("ยา 40", 1)
   Button "Button_12" at 24,16 size 94x40; TextOff 'Back'
      on Press: ActivateScreen("21-30", 0)
   GraphicView "Template_Graphic view_1" at 693,20 size 36x32; Picture "play"
   GraphicView "Template_Graphic view_2" at 27,19 size 36x32; Picture "fast-backward"
   GraphicView "Template_Graphic view_3" at 38,127 size 120x112; Picture "Picture31"
   GraphicView "Template_Graphic view_4" at 190,128 size 120x112; Picture "Picture32"
   GraphicView "Template_Graphic view_5" at 340,128 size 120x112; Picture "Picture33"
   GraphicView "Template_Graphic view_6" at 493,128 size 120x112; Picture "Picture34"
   GraphicView "Template_Graphic view_7" at 644,128 size 120x112; Picture "Picture35"
   GraphicView "Template_Graphic view_8" at 37,302 size 120x112; Picture "Picture36"
   GraphicView "Template_Graphic view_9" at 189,303 size 120x112; Picture "Picture37"
   GraphicView "Template_Graphic view_10" at 339,303 size 120x112; Picture "Picture38"
   GraphicView "Template_Graphic view_11" at 492,303 size 120x112; Picture "Picture39"
   GraphicView "Template_Graphic view_12" at 643,303 size 120x112; Picture "Picture40"
   TextField "Template_Text field_2" at 201,80 size 20x32; Text '4'

screen "41-50" 800x480, template "Template_2"
   Button "Button_1" at 38,239 size 120x40; TextOff 'Magnesium sulfate'
      on Click: ActivateScreen("4_ORDER", 0); SetTag("Selected_URL", 'file:///C:/ASRS_Video/clip41.html')
      on Activate: SetTag("Selected_Medicine", 41)
      on Release: SetTag("ยา 41", 0)
      on Press: SetTag("ยา 41", 1)
   Button "Button_9" at 688,16 size 96x40; TextOff 'Next'
      on Press: ActivateScreen("51-60", 0)
   Button "Button_10" at 38,415 size 120x40; TextOff 'Insulin regular'
      on Click: ActivateScreen("4_ORDER", 0); SetTag("Selected_URL", 'file:///C:/ASRS_Video/clip46.html')
      on Activate: SetTag("Selected_Medicine", 46)
      on Release: SetTag("ยา 46", 0)
      on Press: SetTag("ยา 46", 1)
   Button "Button_2" at 189,240 size 120x40; TextOff 'Calcium gluconate'
      on Click: ActivateScreen("4_ORDER", 0); SetTag("Selected_URL", 'file:///C:/ASRS_Video/clip42.html')
      on Activate: SetTag("Selected_Medicine", 42)
      on Release: SetTag("ยา 42", 0)
      on Press: SetTag("ยา 42", 1)
   Button "Button_3" at 190,415 size 120x40; TextOff 'Glucagon'
      on Click: ActivateScreen("4_ORDER", 0); SetTag("Selected_URL", 'file:///C:/ASRS_Video/clip47.html')
      on Activate: SetTag("Selected_Medicine", 47)
      on Release: SetTag("ยา 47", 0)
      on Press: SetTag("ยา 47", 1)
   Button "Button_4" at 340,240 size 120x40; TextOff 'Sodium bicarbonate'
      on Click: ActivateScreen("4_ORDER", 0); SetTag("Selected_URL", 'file:///C:/ASRS_Video/clip43.html')
      on Activate: SetTag("Selected_Medicine", 43)
      on Release: SetTag("ยา 43", 0)
      on Press: SetTag("ยา 43", 1)
   Button "Button_5" at 340,416 size 120x40; TextOff 'Hydrocortisone'
      on Click: ActivateScreen("4_ORDER", 0); SetTag("Selected_URL", 'file:///C:/ASRS_Video/clip48.html')
      on Activate: SetTag("Selected_Medicine", 48)
      on Release: SetTag("ยา 48", 0)
      on Press: SetTag("ยา 48", 1)
   Button "Button_6" at 494,416 size 120x40; TextOff 'Dexamethasone'
      on Click: ActivateScreen("4_ORDER", 0); SetTag("Selected_URL", 'file:///C:/ASRS_Video/clip49.html')
      on Activate: SetTag("Selected_Medicine", 49)
      on Release: SetTag("ยา 49", 0)
      on Press: SetTag("ยา 49", 1)
   Button "Button_7" at 492,240 size 120x40; TextOff 'Potassium chloride'
      on Click: ActivateScreen("4_ORDER", 0); SetTag("Selected_URL", 'file:///C:/ASRS_Video/clip44.html')
      on Activate: SetTag("Selected_Medicine", 44)
      on Release: SetTag("ยา 44", 0)
      on Press: SetTag("ยา 44", 1)
   Button "Button_8" at 644,240 size 120x40; TextOff 'Dextrose 50%'
      on Click: ActivateScreen("4_ORDER", 0); SetTag("Selected_URL", 'file:///C:/ASRS_Video/clip45.html')
      on Activate: SetTag("Selected_Medicine", 45)
      on Release: SetTag("ยา 45", 0)
      on Press: SetTag("ยา 45", 1)
   Button "Button_11" at 645,416 size 120x40; TextOff 'Diphenhydramine'
      on Click: ActivateScreen("4_ORDER", 0); SetTag("Selected_URL", 'file:///C:/ASRS_Video/clip50.html')
      on Activate: SetTag("Selected_Medicine", 50)
      on Release: SetTag("ยา 50", 0)
      on Press: SetTag("ยา 50", 1)
   Button "Button_12" at 24,16 size 94x40; TextOff 'Back'
      on Press: ActivateScreen("31-40", 0)
   GraphicView "Template_Graphic view_1" at 693,20 size 36x32; Picture "play"
   GraphicView "Template_Graphic view_2" at 27,19 size 36x32; Picture "fast-backward"
   GraphicView "Template_Graphic view_3" at 38,127 size 120x112; Picture "Picture41"
   GraphicView "Template_Graphic view_4" at 190,128 size 120x112; Picture "Picture42"
   GraphicView "Template_Graphic view_5" at 340,128 size 120x112; Picture "Picture43"
   GraphicView "Template_Graphic view_6" at 493,128 size 120x112; Picture "Picture44"
   GraphicView "Template_Graphic view_7" at 644,128 size 120x112; Picture "Picture45"
   GraphicView "Template_Graphic view_8" at 37,302 size 120x112; Picture "Picture46"
   GraphicView "Template_Graphic view_9" at 189,303 size 120x112; Picture "Picture47"
   GraphicView "Template_Graphic view_10" at 339,303 size 120x112; Picture "Picture48"
   GraphicView "Template_Graphic view_11" at 492,303 size 120x112; Picture "Picture49"
   GraphicView "Template_Graphic view_12" at 643,303 size 120x112; Picture "Picture50"
   TextField "Template_Text field_2" at 201,80 size 20x32; Text '5'

screen "51-60" 800x480, template "Template_2"
   Button "Button_1" at 38,239 size 120x40; TextOff 'Chlorpheniramine'
      on Click: ActivateScreen("4_ORDER", 0); SetTag("Selected_URL", 'file:///C:/ASRS_Video/clip51.html')
      on Activate: SetTag("Selected_Medicine", 51)
      on Release: SetTag("ยา 51", 0)
      on Press: SetTag("ยา 51", 1)
   Button "Button_9" at 688,16 size 96x40; TextOff 'Next'
      on Press: ActivateScreen("61-70", 0)
   Button "Button_10" at 38,415 size 120x40; TextOff 'Mannitol'
      on Click: ActivateScreen("4_ORDER", 0); SetTag("Selected_URL", 'file:///C:/ASRS_Video/clip56.html')
      on Activate: SetTag("Selected_Medicine", 56)
      on Release: SetTag("ยา 56", 0)
      on Press: SetTag("ยา 56", 1)
   Button "Button_2" at 189,240 size 120x40; TextOff 'Salbutamol'
      on Click: ActivateScreen("4_ORDER", 0); SetTag("Selected_URL", 'file:///C:/ASRS_Video/clip52.html')
      on Activate: SetTag("Selected_Medicine", 52)
      on Release: SetTag("ยา 52", 0)
      on Press: SetTag("ยา 52", 1)
   Button "Button_3" at 190,415 size 120x40; TextOff 'Acetazolamide'
      on Click: ActivateScreen("4_ORDER", 0); SetTag("Selected_URL", 'file:///C:/ASRS_Video/clip57.html')
      on Activate: SetTag("Selected_Medicine", 57)
      on Release: SetTag("ยา 57", 0)
      on Press: SetTag("ยา 57", 1)
   Button "Button_4" at 340,240 size 120x40; TextOff 'Ipratropium bromide'
      on Click: ActivateScreen("4_ORDER", 0); SetTag("Selected_URL", 'file:///C:/ASRS_Video/clip53.html')
      on Activate: SetTag("Selected_Medicine", 53)
      on Release: SetTag("ยา 53", 0)
      on Press: SetTag("ยา 53", 1)
   Button "Button_5" at 340,416 size 120x40; TextOff 'Tranexamic acid'
      on Click: ActivateScreen("4_ORDER", 0); SetTag("Selected_URL", 'file:///C:/ASRS_Video/clip58.html')
      on Activate: SetTag("Selected_Medicine", 58)
      on Release: SetTag("ยา 58", 0)
      on Press: SetTag("ยา 58", 1)
   Button "Button_6" at 492,416 size 120x40; TextOff 'Vitamin K'
      on Click: ActivateScreen("4_ORDER", 0); SetTag("Selected_URL", 'file:///C:/ASRS_Video/clip59.html')
      on Activate: SetTag("Selected_Medicine", 59)
      on Release: SetTag("ยา 59", 0)
      on Press: SetTag("ยา 59", 1)
   Button "Button_7" at 492,240 size 120x40; TextOff 'Aminophylline'
      on Click: ActivateScreen("4_ORDER", 0); SetTag("Selected_URL", 'file:///C:/ASRS_Video/clip54.html')
      on Activate: SetTag("Selected_Medicine", 54)
      on Release: SetTag("ยา 54", 0)
      on Press: SetTag("ยา 54", 1)
   Button "Button_8" at 644,240 size 120x40; TextOff 'Furosemide'
      on Click: ActivateScreen("4_ORDER", 0); SetTag("Selected_URL", 'file:///C:/ASRS_Video/clip55.html')
      on Activate: SetTag("Selected_Medicine", 55)
      on Release: SetTag("ยา 55", 0)
      on Press: SetTag("ยา 55", 1)
   Button "Button_11" at 645,416 size 120x40; TextOff 'Protamine sulfate'
      on Click: ActivateScreen("4_ORDER", 0); SetTag("Selected_URL", 'file:///C:/ASRS_Video/clip60.html')
      on Activate: SetTag("Selected_Medicine", 60)
      on Release: SetTag("ยา 60", 0)
      on Press: SetTag("ยา 60", 1)
   Button "Button_12" at 24,16 size 94x40; TextOff 'Back'
      on Press: ActivateScreen("41-50", 0)
   GraphicView "Template_Graphic view_1" at 693,20 size 36x32; Picture "play"
   GraphicView "Template_Graphic view_2" at 27,19 size 36x32; Picture "fast-backward"
   GraphicView "Template_Graphic view_3" at 38,127 size 120x112; Picture "Picture51"
   GraphicView "Template_Graphic view_4" at 190,128 size 120x112; Picture "Picture52"
   GraphicView "Template_Graphic view_5" at 340,128 size 120x112; Picture "Picture53"
   GraphicView "Template_Graphic view_6" at 493,128 size 120x112; Picture "Picture54"
   GraphicView "Template_Graphic view_7" at 644,128 size 120x112; Picture "Picture55"
   GraphicView "Template_Graphic view_8" at 37,302 size 120x112; Picture "Picture56"
   GraphicView "Template_Graphic view_9" at 189,303 size 120x112; Picture "Picture57"
   GraphicView "Template_Graphic view_10" at 339,303 size 120x112; Picture "Picture58"
   GraphicView "Template_Graphic view_11" at 492,303 size 120x112; Picture "Picture59"
   GraphicView "Template_Graphic view_12" at 643,303 size 120x112; Picture "Picture60"
   TextField "Template_Text field_2" at 201,80 size 20x32; Text '6'

screen "61-70" 800x480, template "Template_2"
   Button "Button_1" at 28,239 size 120x40; TextOff 'Naloxone'
      on Click: ActivateScreen("4_ORDER", 0); SetTag("Selected_URL", 'file:///C:/ASRS_Video/clip61.html')
      on Activate: SetTag("Selected_Medicine", 61)
      on Release: SetTag("ยา 61", 0)
      on Press: SetTag("ยา 61", 1)
   Button "Button_9" at 688,16 size 96x40; TextOff 'Next'
      on Press: ActivateScreen("71-80", 0)
   Button "Button_10" at 28,415 size 120x40; TextOff 'Pralidoxime'
      on Click: ActivateScreen("4_ORDER", 0); SetTag("Selected_URL", 'file:///C:/ASRS_Video/clip66.html')
      on Activate: SetTag("Selected_Medicine", 66)
      on Release: SetTag("ยา 66", 0)
      on Press: SetTag("ยา 66", 1)
   Button "Button_2" at 182,240 size 120x40; TextOff 'Flumazenil'
      on Click: ActivateScreen("4_ORDER", 0); SetTag("Selected_URL", 'file:///C:/ASRS_Video/clip62.html')
      on Activate: SetTag("Selected_Medicine", 62)
      on Release: SetTag("ยา 62", 0)
      on Press: SetTag("ยา 62", 1)
   Button "Button_3" at 183,415 size 120x40; TextOff 'Atropine'
      on Click: ActivateScreen("4_ORDER", 0); SetTag("Selected_URL", 'file:///C:/ASRS_Video/clip67.html')
      on Activate: SetTag("Selected_Medicine", 67)
      on Release: SetTag("ยา 67", 0)
      on Press: SetTag("ยา 67", 1)
   Button "Button_4" at 333,240 size 120x40; TextOff 'Activated charcoal'
      on Click: ActivateScreen("4_ORDER", 0); SetTag("Selected_URL", 'file:///C:/ASRS_Video/clip63.html')
      on Activate: SetTag("Selected_Medicine", 63)
      on Release: SetTag("ยา 63", 0)
      on Press: SetTag("ยา 63", 1)
   Button "Button_5" at 333,416 size 120x40; TextOff 'Methylene blue'
      on Click: ActivateScreen("4_ORDER", 0); SetTag("Selected_URL", 'file:///C:/ASRS_Video/clip68.html')
      on Activate: SetTag("Selected_Medicine", 68)
      on Release: SetTag("ยา 68", 0)
      on Press: SetTag("ยา 68", 1)
   Button "Button_6" at 485,416 size 120x40; TextOff 'Succimer'
      on Click: ActivateScreen("4_ORDER", 0); SetTag("Selected_URL", 'file:///C:/ASRS_Video/clip69.html')
      on Activate: SetTag("Selected_Medicine", 69)
      on Release: SetTag("ยา 69", 0)
      on Press: SetTag("ยา 69", 1)
   Button "Button_7" at 485,240 size 120x40; TextOff 'Acetylcysteine'
      on Click: ActivateScreen("4_ORDER", 0); SetTag("Selected_URL", 'file:///C:/ASRS_Video/clip64.html')
      on Activate: SetTag("Selected_Medicine", 64)
      on Release: SetTag("ยา 64", 0)
      on Press: SetTag("ยา 64", 1)
   Button "Button_8" at 637,240 size 120x40; TextOff 'Deferoxamine'
      on Click: ActivateScreen("4_ORDER", 0); SetTag("Selected_URL", 'file:///C:/ASRS_Video/clip65.html')
      on Activate: SetTag("Selected_Medicine", 65)
      on Release: SetTag("ยา 65", 0)
      on Press: SetTag("ยา 65", 1)
   Button "Button_11" at 638,416 size 120x40; TextOff 'Digoxin immune fab'
      on Click: ActivateScreen("4_ORDER", 0); SetTag("Selected_URL", 'file:///C:/ASRS_Video/clip70.html')
      on Activate: SetTag("Selected_Medicine", 70)
      on Release: SetTag("ยา 70", 0)
      on Press: SetTag("ยา 70", 1)
   Button "Button_12" at 24,16 size 94x40; TextOff 'Back'
      on Press: ActivateScreen("51-60", 0)
   GraphicView "Template_Graphic view_1" at 693,20 size 36x32; Picture "play"
   GraphicView "Template_Graphic view_2" at 27,19 size 36x32; Picture "fast-backward"
   GraphicView "Template_Graphic view_3" at 29,127 size 120x112; Picture "Picture61"
   GraphicView "Template_Graphic view_4" at 186,128 size 120x112; Picture "Picture62"
   GraphicView "Template_Graphic view_5" at 331,128 size 120x112; Picture "Picture63"
   GraphicView "Template_Graphic view_6" at 487,128 size 120x112; Picture "Picture64"
   GraphicView "Template_Graphic view_7" at 637,128 size 120x112; Picture "Picture65"
   GraphicView "Template_Graphic view_8" at 29,302 size 120x112; Picture "Picture66"
   GraphicView "Template_Graphic view_9" at 181,303 size 120x104; Picture "Picture67"
   GraphicView "Template_Graphic view_10" at 330,303 size 120x112; Picture "Picture68"
   GraphicView "Template_Graphic view_11" at 481,303 size 120x112; Picture "Picture69"
   GraphicView "Template_Graphic view_12" at 634,303 size 120x104; Picture "Picture70"
   TextField "Template_Text field_2" at 201,80 size 20x32; Text '7'

screen "71-80" 800x480, template "Template_2"
   Button "Button_1" at 38,239 size 120x40; TextOff 'Fomepizole'
      on Click: ActivateScreen("4_ORDER", 0); SetTag("Selected_URL", 'file:///C:/ASRS_Video/clip71.html')
      on Activate: SetTag("Selected_Medicine", 71)
      on Release: SetTag("ยา 71", 0)
      on Press: SetTag("ยา 71", 1)
   Button "Button_10" at 38,415 size 120x40; TextOff 'Normal saline'
      on Click: ActivateScreen("4_ORDER", 0); SetTag("Selected_URL", 'file:///C:/ASRS_Video/clip76.html')
      on Activate: SetTag("Selected_Medicine", 76)
      on Release: SetTag("ยา 76", 0)
      on Press: SetTag("ยา 76", 1)
   Button "Button_2" at 189,240 size 120x40; TextOff 'Antivenom green pit viper'
      on Click: ActivateScreen("4_ORDER", 0); SetTag("Selected_URL", 'file:///C:/ASRS_Video/clip72.html')
      on Activate: SetTag("Selected_Medicine", 72)
      on Release: SetTag("ยา 72", 0)
      on Press: SetTag("ยา 72", 1)
   Button "Button_3" at 190,415 size 120x40; TextOff 'Heparin'
      on Click: ActivateScreen("4_ORDER", 0); SetTag("Selected_URL", 'file:///C:/ASRS_Video/clip77.html')
      on Activate: SetTag("Selected_Medicine", 77)
      on Release: SetTag("ยา 77", 0)
      on Press: SetTag("ยา 77", 1)
   Button "Button_4" at 340,240 size 120x40; TextOff 'Rabies immunoglobulin'
      on Click: ActivateScreen("4_ORDER", 0); SetTag("Selected_URL", 'file:///C:/ASRS_Video/clip73.html')
      on Activate: SetTag("Selected_Medicine", 73)
      on Release: SetTag("ยา 73", 0)
      on Press: SetTag("ยา 73", 1)
   Button "Button_5" at 340,416 size 120x40; TextOff 'Enoxaparin'
      on Click: ActivateScreen("4_ORDER", 0); SetTag("Selected_URL", 'file:///C:/ASRS_Video/clip78.html')
      on Activate: SetTag("Selected_Medicine", 78)
      on Release: SetTag("ยา 78", 0)
      on Press: SetTag("ยา 78", 1)
   Button "Button_6" at 492,416 size 120x40; TextOff 'Alteplase'
      on Click: ActivateScreen("4_ORDER", 0); SetTag("Selected_URL", 'file:///C:/ASRS_Video/clip79.html')
      on Activate: SetTag("Selected_Medicine", 79)
      on Release: SetTag("ยา 79", 0)
      on Press: SetTag("ยา 79", 1)
   Button "Button_7" at 492,240 size 120x40; TextOff 'Tetanus immunoglobulin'
      on Click: ActivateScreen("4_ORDER", 0); SetTag("Selected_URL", 'file:///C:/ASRS_Video/clip74.html')
      on Activate: SetTag("Selected_Medicine", 74)
      on Release: SetTag("ยา 74", 0)
      on Press: SetTag("ยา 74", 1)
   Button "Button_8" at 644,240 size 120x40; TextOff 'Human albumin'
      on Click: ActivateScreen("4_ORDER", 0); SetTag("Selected_URL", 'file:///C:/ASRS_Video/clip75.html')
      on Activate: SetTag("Selected_Medicine", 75)
      on Release: SetTag("ยา 75", 0)
      on Press: SetTag("ยา 75", 1)
   Button "Button_11" at 645,416 size 120x40; TextOff 'Streptokinase'
      on Click: ActivateScreen("4_ORDER", 0); SetTag("Selected_URL", 'file:///C:/ASRS_Video/clip80.html')
      on Activate: SetTag("Selected_Medicine", 80)
      on Release: SetTag("ยา 80", 0)
      on Press: SetTag("ยา 80", 1)
   Button "Button_12" at 24,16 size 94x40; TextOff 'Back'
      on Press: ActivateScreen("61-70", 0)
   Button "Button_9" at 688,16 size 96x40; TextOff 'Next'
      on Press: ActivateScreen("81-90", 0)
   GraphicView "Template_Graphic view_2" at 27,19 size 36x32; Picture "fast-backward"
   GraphicView "Template_Graphic view_1" at 693,20 size 36x32; Picture "play"
   GraphicView "Template_Graphic view_3" at 37,128 size 120x104; Picture "Picture71"
   GraphicView "Template_Graphic view_4" at 191,129 size 120x104; Picture "Picture72"
   GraphicView "Template_Graphic view_5" at 339,129 size 120x104; Picture "Picture73"
   GraphicView "Template_Graphic view_6" at 493,129 size 120x104; Picture "Picture74"
   GraphicView "Template_Graphic view_7" at 645,129 size 120x112; Picture "Picture75"
   GraphicView "Template_Graphic view_8" at 35,303 size 120x112; Picture "Picture76"
   GraphicView "Template_Graphic view_9" at 189,304 size 120x112; Picture "Picture77"
   GraphicView "Template_Graphic view_10" at 338,304 size 120x104; Picture "Picture78"
   GraphicView "Template_Graphic view_11" at 497,304 size 120x112; Picture "Picture79"
   GraphicView "Template_Graphic view_12" at 645,304 size 120x112; Picture "Picture80"
   TextField "Template_Text field_2" at 201,80 size 20x32; Text '8'

screen "81-90" 800x480, template "Template_2"
   Button "Button_1" at 38,239 size 120x40; TextOff 'Urokinase'
      on Click: ActivateScreen("4_ORDER", 0); SetTag("Selected_URL", 'file:///C:/ASRS_Video/clip81.html')
      on Activate: SetTag("Selected_Medicine", 81)
      on Release: SetTag("ยา 81", 0)
      on Press: SetTag("ยา 81", 1)
   Button "Button_10" at 38,415 size 120x40; TextOff 'Haloperidol'
      on Click: ActivateScreen("4_ORDER", 0); SetTag("Selected_URL", 'file:///C:/ASRS_Video/clip86.html')
      on Activate: SetTag("Selected_Medicine", 86)
      on Release: SetTag("ยา 86", 0)
      on Press: SetTag("ยา 86", 1)
   Button "Button_2" at 189,240 size 120x40; TextOff 'Iohexol'
      on Click: ActivateScreen("4_ORDER", 0); SetTag("Selected_URL", 'file:///C:/ASRS_Video/clip82.html')
      on Activate: SetTag("Selected_Medicine", 82)
      on Release: SetTag("ยา 82", 0)
      on Press: SetTag("ยา 82", 1)
   Button "Button_3" at 190,415 size 120x40; TextOff 'Olanzapine'
      on Click: ActivateScreen("4_ORDER", 0); SetTag("Selected_URL", 'file:///C:/ASRS_Video/clip87.html')
      on Activate: SetTag("Selected_Medicine", 87)
      on Release: SetTag("ยา 87", 0)
      on Press: SetTag("ยา 87", 1)
   Button "Button_4" at 340,240 size 120x40; TextOff 'Iopamidol'
      on Click: ActivateScreen("4_ORDER", 0); SetTag("Selected_URL", 'file:///C:/ASRS_Video/clip83.html')
      on Activate: SetTag("Selected_Medicine", 83)
      on Release: SetTag("ยา 83", 0)
      on Press: SetTag("ยา 83", 1)
   Button "Button_5" at 340,416 size 120x40; TextOff 'Levetiracetam'
      on Click: ActivateScreen("4_ORDER", 0); SetTag("Selected_URL", 'file:///C:/ASRS_Video/clip88.html')
      on Activate: SetTag("Selected_Medicine", 88)
      on Release: SetTag("ยา 88", 0)
      on Press: SetTag("ยา 88", 1)
   Button "Button_6" at 492,416 size 120x40; TextOff 'Phenytoin'
      on Click: ActivateScreen("4_ORDER", 0); SetTag("Selected_URL", 'file:///C:/ASRS_Video/clip89.html')
      on Activate: SetTag("Selected_Medicine", 89)
      on Release: SetTag("ยา 89", 0)
      on Press: SetTag("ยา 89", 1)
   Button "Button_7" at 492,240 size 120x40; TextOff 'Iodixanol'
      on Click: ActivateScreen("4_ORDER", 0); SetTag("Selected_URL", 'file:///C:/ASRS_Video/clip84.html')
      on Activate: SetTag("Selected_Medicine", 84)
      on Release: SetTag("ยา 84", 0)
      on Press: SetTag("ยา 84", 1)
   Button "Button_8" at 644,240 size 120x40; TextOff 'Gadopentetate dimeglumine'
      on Click: ActivateScreen("4_ORDER", 0); SetTag("Selected_URL", 'file:///C:/ASRS_Video/clip85.html')
      on Activate: SetTag("Selected_Medicine", 85)
      on Release: SetTag("ยา 85", 0)
      on Press: SetTag("ยา 85", 1)
   Button "Button_11" at 645,416 size 120x40; TextOff 'Sodium valproate'
      on Click: ActivateScreen("4_ORDER", 0); SetTag("Selected_URL", 'file:///C:/ASRS_Video/clip90.html')
      on Activate: SetTag("Selected_Medicine", 90)
      on Release: SetTag("ยา 90", 0)
      on Press: SetTag("ยา 90", 1)
   Button "Button_12" at 24,16 size 94x40; TextOff 'Back'
      on Press: ActivateScreen("71-80", 0)
   Button "Button_9" at 688,16 size 96x40; TextOff 'Next'
      on Press: ActivateScreen("91-100", 0)
   GraphicView "Template_Graphic view_2" at 27,19 size 36x32; Picture "fast-backward"
   GraphicView "Template_Graphic view_1" at 693,20 size 36x32; Picture "play"
   GraphicView "Template_Graphic view_3" at 37,128 size 120x104; Picture "Picture81"
   GraphicView "Template_Graphic view_4" at 191,129 size 120x104; Picture "Picture82"
   GraphicView "Template_Graphic view_5" at 339,129 size 120x104; Picture "Picture83"
   GraphicView "Template_Graphic view_6" at 493,129 size 120x104; Picture "Picture84"
   GraphicView "Template_Graphic view_7" at 645,129 size 120x112; Picture "Picture85"
   GraphicView "Template_Graphic view_8" at 38,305 size 120x104; Picture "Picture86"
   GraphicView "Template_Graphic view_9" at 189,304 size 120x112; Picture "Picture87"
   GraphicView "Template_Graphic view_10" at 338,304 size 120x112; Picture "Picture88"
   GraphicView "Template_Graphic view_11" at 497,304 size 120x112; Picture "Picture89"
   GraphicView "Template_Graphic view_12" at 645,304 size 120x112; Picture "Picture90"
   TextField "Template_Text field_2" at 201,80 size 20x32; Text '9'

screen "91-100" 800x480, template "Template_2"
   Button "Button_1" at 38,239 size 120x40; TextOff 'Carbamazepine'
      on Click: ActivateScreen("4_ORDER", 0); SetTag("Selected_URL", 'file:///C:/ASRS_Video/clip91.html')
      on Activate: SetTag("Selected_Medicine", 91)
      on Release: SetTag("ยา 91", 0)
      on Press: SetTag("ยา 91", 1)
   Button "Button_10" at 38,415 size 120x40; TextOff 'Metoclopramide'
      on Click: ActivateScreen("4_ORDER", 0); SetTag("Selected_URL", 'file:///C:/ASRS_Video/clip96.html')
      on Activate: SetTag("Selected_Medicine", 1)
      on Release: SetTag("ยา 96", 0)
      on Press: SetTag("ยา 96", 1)
   Button "Button_2" at 189,240 size 120x40; TextOff 'Phenobarbital'
      on Click: ActivateScreen("4_ORDER", 0); SetTag("Selected_URL", 'file:///C:/ASRS_Video/clip92.html')
      on Activate: SetTag("Selected_Medicine", 92)
      on Release: SetTag("ยา 92", 0)
      on Press: SetTag("ยา 92", 1)
   Button "Button_3" at 190,415 size 120x40; TextOff 'Granisetron'
      on Click: ActivateScreen("4_ORDER", 0); SetTag("Selected_URL", 'file:///C:/ASRS_Video/clip97.html')
      on Activate: SetTag("Selected_Medicine", 97)
      on Release: SetTag("ยา 97", 0)
      on Press: SetTag("ยา 97", 1)
   Button "Button_4" at 340,240 size 120x40; TextOff 'Ketorolac'
      on Click: ActivateScreen("4_ORDER", 0); SetTag("Selected_URL", 'file:///C:/ASRS_Video/clip93.html')
      on Activate: SetTag("Selected_Medicine", 93)
      on Release: SetTag("ยา 93", 0)
      on Press: SetTag("ยา 93", 1)
   Button "Button_5" at 340,416 size 120x40; TextOff 'Sugammadex'
      on Click: ActivateScreen("4_ORDER", 0); SetTag("Selected_URL", 'file:///C:/ASRS_Video/clip98.html')
      on Activate: SetTag("Selected_Medicine", 98)
      on Release: SetTag("ยา 98", 0)
      on Press: SetTag("ยา 98", 1)
   Button "Button_6" at 492,416 size 120x40; TextOff 'Hydrocolloid dressing'
      on Click: ActivateScreen("4_ORDER", 0); SetTag("Selected_URL", 'file:///C:/ASRS_Video/clip99.html')
      on Activate: SetTag("Selected_Medicine", 99)
      on Release: SetTag("ยา 99", 0)
      on Press: SetTag("ยา 99", 1)
   Button "Button_7" at 492,240 size 120x40; TextOff 'Parecoxib'
      on Click: ActivateScreen("4_ORDER", 0); SetTag("Selected_URL", 'file:///C:/ASRS_Video/clip94.html')
      on Activate: SetTag("Selected_Medicine", 94)
      on Release: SetTag("ยา 94", 0)
      on Press: SetTag("ยา 94", 1)
   Button "Button_8" at 644,240 size 120x40; TextOff 'Ondansetron'
      on Click: ActivateScreen("4_ORDER", 0); SetTag("Selected_URL", 'file:///C:/ASRS_Video/clip95.html')
      on Activate: SetTag("Selected_Medicine", 95)
      on Release: SetTag("ยา 95", 0)
      on Press: SetTag("ยา 95", 1)
   Button "Button_11" at 645,416 size 120x40; TextOff 'Paraffin gauze dressing'
      on Click: ActivateScreen("4_ORDER", 0); SetTag("Selected_URL", 'file:///C:/ASRS_Video/clip100.html')
      on Activate: SetTag("Selected_Medicine", 100)
      on Release: SetTag("ยา 100", 0)
      on Press: SetTag("ยา 100", 1)
   Button "Button_12" at 24,16 size 94x40; TextOff 'Back'
      on Press: ActivateScreen("81-90", 0)
   GraphicView "Template_Graphic view_2" at 27,19 size 36x32; Picture "fast-backward"
   GraphicView "Template_Graphic view_3" at 37,128 size 120x104; Picture "Picture91"
   GraphicView "Template_Graphic view_4" at 191,129 size 120x104; Picture "Picture92"
   GraphicView "Template_Graphic view_5" at 339,129 size 120x104; Picture "Picture93"
   GraphicView "Template_Graphic view_6" at 493,129 size 120x104; Picture "Picture94"
   GraphicView "Template_Graphic view_7" at 645,129 size 120x104; Picture "Picture95"
   GraphicView "Template_Graphic view_8" at 38,305 size 120x104; Picture "Picture96"
   GraphicView "Template_Graphic view_9" at 189,304 size 120x112; Picture "Picture97"
   GraphicView "Template_Graphic view_10" at 351,307 size 96x104; Picture "Picture98"
   GraphicView "Template_Graphic view_11" at 497,304 size 120x112; Picture "Picture99"
   GraphicView "Template_Graphic view_12" at 645,304 size 120x104; Picture "Picture100"
   TextField "Template_Text field_2" at 201,80 size 36x32; Text '10'

screen "1" 800x480, template "Template_2"
   Button "Button_1" at 40,240 size 120x40; TextOff 'Omeprazole'
      on Click: ActivateScreen("4_ORDER", 0); SetTag("Selected_URL", 'file:///C:/ASRS_Video/clip101.html')
      on Activate: SetTag("Selected_Medicine", 101)
      on Release: SetTag("ยา 101", 0)
      on Press: SetTag("ยา 101", 1)
   Button "Button_10" at 38,415 size 120x40; TextOff 'Famotidine'
      on Click: ActivateScreen("4_ORDER", 0); SetTag("Selected_URL", 'file:///C:/ASRS_Video/clip106.html')
      on Activate: SetTag("Selected_Medicine", 106)
      on Release: SetTag("ยา 106", 0)
      on Press: SetTag("ยา 106", 1)
   Button "Button_2" at 189,240 size 120x40; TextOff 'Esomeprazole'
      on Click: ActivateScreen("4_ORDER", 0); SetTag("Selected_URL", 'file:///C:/ASRS_Video/clip102.html')
      on Activate: SetTag("Selected_Medicine", 102)
      on Release: SetTag("ยา 102", 0)
      on Press: SetTag("ยา 102", 1)
   Button "Button_3" at 190,415 size 120x40; TextOff 'Cimetidine'
      on Click: ActivateScreen("4_ORDER", 0); SetTag("Selected_URL", 'file:///C:/ASRS_Video/clip107.html')
      on Activate: SetTag("Selected_Medicine", 107)
      on Release: SetTag("ยา 107", 0)
      on Press: SetTag("ยา 107", 1)
   Button "Button_4" at 340,240 size 120x40; TextOff 'Pantoprazole'
      on Click: ActivateScreen("4_ORDER", 0); SetTag("Selected_URL", 'file:///C:/ASRS_Video/clip103.html')
      on Activate: SetTag("Selected_Medicine", 103)
      on Release: SetTag("ยา 103", 0)
      on Press: SetTag("ยา 103", 1)
   Button "Button_5" at 340,416 size 120x40; TextOff 'Sucralfate'
      on Click: ActivateScreen("4_ORDER", 0); SetTag("Selected_URL", 'file:///C:/ASRS_Video/clip108.html')
      on Activate: SetTag("Selected_Medicine", 108)
      on Release: SetTag("ยา 108", 0)
      on Press: SetTag("ยา 108", 1)
   Button "Button_6" at 492,416 size 120x40; TextOff 'Aluminium hydroxide'
      on Click: ActivateScreen("4_ORDER", 0); SetTag("Selected_URL", 'file:///C:/ASRS_Video/clip109.html')
      on Activate: SetTag("Selected_Medicine", 109)
      on Release: SetTag("ยา 109", 0)
      on Press: SetTag("ยา 109", 1)
   Button "Button_7" at 492,240 size 120x40; TextOff 'Lansoprazole'
      on Click: ActivateScreen("4_ORDER", 0); SetTag("Selected_URL", 'file:///C:/ASRS_Video/clip104.html')
      on Activate: SetTag("Selected_Medicine", 104)
      on Release: SetTag("ยา 104", 0)
      on Press: SetTag("ยา 104", 1)
   Button "Button_8" at 644,240 size 120x40; TextOff 'Dexlansoprazole'
      on Click: ActivateScreen("4_ORDER", 0); SetTag("Selected_URL", 'file:///C:/ASRS_Video/clip105.html')
      on Activate: SetTag("Selected_Medicine", 105)
      on Release: SetTag("ยา 105", 0)
      on Press: SetTag("ยา 105", 1)
   Button "Button_11" at 645,416 size 120x40; TextOff 'Magnesium hydroxide'
      on Click: ActivateScreen("4_ORDER", 0); SetTag("Selected_URL", 'file:///C:/ASRS_Video/clip110.html')
      on Activate: SetTag("Selected_Medicine", 110)
      on Release: SetTag("ยา 110", 0)
      on Press: SetTag("ยา 110", 1)
   Button "Button_12" at 688,16 size 96x40; TextOff 'Next'
      on Press: ActivateScreen("2", 0)
   Button "Button_9" at 24,16 size 94x40; TextOff 'Back'
      on Press: ActivateScreen("4_ORDER", 0)
   GraphicView "Template_Graphic view_2" at 693,20 size 36x32; Picture "play"
   GraphicView "Template_Graphic view_1" at 27,19 size 36x32; Picture "fast-backward"
   GraphicView "Template_Graphic view_3" at 37,128 size 120x104; Picture "Picture101"
   GraphicView "Template_Graphic view_4" at 191,129 size 120x104; Picture "Picture102"
   GraphicView "Template_Graphic view_5" at 339,129 size 120x104; Picture "Picture103"
   GraphicView "Template_Graphic view_6" at 493,129 size 120x104; Picture "Picture104"
   GraphicView "Template_Graphic view_7" at 645,129 size 120x104; Picture "Picture105"
   GraphicView "Template_Graphic view_8" at 38,305 size 120x104; Picture "Picture106"
   GraphicView "Template_Graphic view_9" at 189,304 size 120x112; Picture "Picture107"
   GraphicView "Template_Graphic view_10" at 351,307 size 96x104; Picture "Picture108"
   GraphicView "Template_Graphic view_11" at 497,304 size 120x112; Picture "Picture109"
   GraphicView "Template_Graphic view_12" at 645,304 size 120x104; Picture "Picture110"
   TextField "Template_Text field_2" at 201,80 size 20x32; Text '1'

screen "2" 800x480, template "Template_2"
   Button "Button_1" at 38,239 size 120x40; TextOff 'Simethicone'
      on Click: ActivateScreen("4_ORDER", 0); SetTag("Selected_URL", 'file:///C:/ASRS_Video/clip111.html')
      on Activate: SetTag("Selected_Medicine", 111)
      on Release: SetTag("ยา 111", 0)
      on Press: SetTag("ยา 111", 1)
   Button "Button_9" at 688,16 size 96x40; TextOff 'Next'
      on Press: ActivateScreen("3", 0)
   Button "Button_10" at 38,415 size 120x40; TextOff 'Bisacodyl'
      on Click: ActivateScreen("4_ORDER", 0); SetTag("Selected_URL", 'file:///C:/ASRS_Video/clip116.html')
      on Activate: SetTag("Selected_Medicine", 116)
      on Release: SetTag("ยา 116", 0)
      on Press: SetTag("ยา 116", 1)
   Button "Button_2" at 189,240 size 120x40; TextOff 'Domperidone'
      on Click: ActivateScreen("4_ORDER", 0); SetTag("Selected_URL", 'file:///C:/ASRS_Video/clip112.html')
      on Activate: SetTag("Selected_Medicine", 112)
      on Release: SetTag("ยา 112", 0)
      on Press: SetTag("ยา 112", 1)
   Button "Button_3" at 190,415 size 120x40; TextOff 'Lactulose'
      on Click: ActivateScreen("4_ORDER", 0); SetTag("Selected_URL", 'file:///C:/ASRS_Video/clip117.html')
      on Activate: SetTag("Selected_Medicine", 117)
      on Release: SetTag("ยา 117", 0)
      on Press: SetTag("ยา 117", 1)
   Button "Button_4" at 340,240 size 120x40; TextOff 'Metoclopramide'
      on Click: ActivateScreen("4_ORDER", 0); SetTag("Selected_URL", 'file:///C:/ASRS_Video/clip113.html')
      on Activate: SetTag("Selected_Medicine", 113)
      on Release: SetTag("ยา 113", 0)
      on Press: SetTag("ยา 113", 1)
   Button "Button_5" at 340,416 size 120x40; TextOff 'Senna'
      on Click: ActivateScreen("4_ORDER", 0); SetTag("Selected_URL", 'file:///C:/ASRS_Video/clip118.html')
      on Activate: SetTag("Selected_Medicine", 118)
      on Release: SetTag("ยา 118", 0)
      on Press: SetTag("ยา 118", 1)
   Button "Button_6" at 492,416 size 120x40; TextOff 'ORS'
      on Click: ActivateScreen("4_ORDER", 0); SetTag("Selected_URL", 'file:///C:/ASRS_Video/clip119.html')
      on Activate: SetTag("Selected_Medicine", 119)
      on Release: SetTag("ยา 119", 0)
      on Press: SetTag("ยา 119", 1)
   Button "Button_7" at 492,240 size 120x40; TextOff 'Ondansetron'
      on Click: ActivateScreen("4_ORDER", 0); SetTag("Selected_URL", 'file:///C:/ASRS_Video/clip114.html')
      on Activate: SetTag("Selected_Medicine", 114)
      on Release: SetTag("ยา 114", 0)
      on Press: SetTag("ยา 114", 1)
   Button "Button_8" at 644,240 size 120x40; TextOff 'Hyoscine butylbromide'
      on Click: ActivateScreen("4_ORDER", 0); SetTag("Selected_URL", 'file:///C:/ASRS_Video/clip115.html')
      on Activate: SetTag("Selected_Medicine", 115)
      on Release: SetTag("ยา 115", 0)
      on Press: SetTag("ยา 115", 1)
   Button "Button_11" at 645,416 size 120x40; TextOff 'Loperamide'
      on Click: ActivateScreen("4_ORDER", 0); SetTag("Selected_URL", 'file:///C:/ASRS_Video/clip120.html')
      on Activate: SetTag("Selected_Medicine", 120)
      on Release: SetTag("ยา 120", 0)
      on Press: SetTag("ยา 120", 1)
   Button "Button_12" at 24,16 size 94x40; TextOff 'Back'
      on Press: ActivateScreen("1", 0)
   GraphicView "Template_Graphic view_1" at 693,20 size 36x32; Picture "play"
   GraphicView "Template_Graphic view_2" at 27,19 size 36x32; Picture "fast-backward"
   GraphicView "Template_Graphic view_3" at 37,128 size 120x104; Picture "Picture111"
   GraphicView "Template_Graphic view_4" at 191,129 size 120x104; Picture "Picture112"
   GraphicView "Template_Graphic view_5" at 339,129 size 120x104; Picture "Picture113"
   GraphicView "Template_Graphic view_6" at 493,129 size 120x104; Picture "Picture114"
   GraphicView "Template_Graphic view_7" at 645,129 size 120x104; Picture "Picture115"
   GraphicView "Template_Graphic view_8" at 38,305 size 120x104; Picture "Picture116"
   GraphicView "Template_Graphic view_9" at 189,304 size 120x104; Picture "Picture117"
   GraphicView "Template_Graphic view_10" at 351,307 size 96x104; Picture "Picture118"
   GraphicView "Template_Graphic view_11" at 497,304 size 120x112; Picture "Picture119"
   GraphicView "Template_Graphic view_12" at 645,304 size 120x104; Picture "Picture120"
   TextField "Template_Text field_2" at 201,80 size 20x32; Text '2'

screen "3" 800x480, template "Template_2"
   Button "Button_1" at 38,239 size 120x40; TextOff 'Amlodipine'
      on Click: ActivateScreen("4_ORDER", 0); SetTag("Selected_URL", 'file:///C:/ASRS_Video/clip121.html')
      on Activate: SetTag("Selected_Medicine", 121)
      on Release: SetTag("ยา 121", 0)
      on Press: SetTag("ยา 121", 1)
   Button "Button_9" at 688,16 size 96x40; TextOff 'Next'
      on Press: ActivateScreen("4", 0)
   Button "Button_10" at 38,415 size 120x40; TextOff 'Hydrochlorothiazide'
      on Click: ActivateScreen("4_ORDER", 0); SetTag("Selected_URL", 'file:///C:/ASRS_Video/clip126.html')
      on Activate: SetTag("Selected_Medicine", 126)
      on Release: SetTag("ยา 126", 0)
      on Press: SetTag("ยา 126", 1)
   Button "Button_2" at 189,240 size 120x40; TextOff 'Losartan'
      on Click: ActivateScreen("4_ORDER", 0); SetTag("Selected_URL", 'file:///C:/ASRS_Video/clip122.html')
      on Activate: SetTag("Selected_Medicine", 122)
      on Release: SetTag("ยา 122", 0)
      on Press: SetTag("ยา 122", 1)
   Button "Button_3" at 190,415 size 120x40; TextOff 'Furosemide'
      on Click: ActivateScreen("4_ORDER", 0); SetTag("Selected_URL", 'file:///C:/ASRS_Video/clip127.html')
      on Activate: SetTag("Selected_Medicine", 127)
      on Release: SetTag("ยา 127", 0)
      on Press: SetTag("ยา 127", 1)
   Button "Button_4" at 340,240 size 120x40; TextOff 'Enalapril'
      on Click: ActivateScreen("4_ORDER", 0); SetTag("Selected_URL", 'file:///C:/ASRS_Video/clip123.html')
      on Activate: SetTag("Selected_Medicine", 123)
      on Release: SetTag("ยา 123", 0)
      on Press: SetTag("ยา 123", 1)
   Button "Button_5" at 340,416 size 120x40; TextOff 'Spironolactone'
      on Click: ActivateScreen("4_ORDER", 0); SetTag("Selected_URL", 'file:///C:/ASRS_Video/clip128.html')
      on Activate: SetTag("Selected_Medicine", 128)
      on Release: SetTag("ยา 128", 0)
      on Press: SetTag("ยา 128", 1)
   Button "Button_6" at 492,416 size 120x40; TextOff 'Atenolol'
      on Click: ActivateScreen("4_ORDER", 0); SetTag("Selected_URL", 'file:///C:/ASRS_Video/clip129.html')
      on Activate: SetTag("Selected_Medicine", 129)
      on Release: SetTag("ยา 129", 0)
      on Press: SetTag("ยา 129", 1)
   Button "Button_7" at 492,240 size 120x40; TextOff 'Captopril'
      on Click: ActivateScreen("4_ORDER", 0); SetTag("Selected_URL", 'file:///C:/ASRS_Video/clip124.html')
      on Activate: SetTag("Selected_Medicine", 124)
      on Release: SetTag("ยา 124", 0)
      on Press: SetTag("ยา 124", 1)
   Button "Button_8" at 644,240 size 120x40; TextOff 'Lisinopril'
      on Click: ActivateScreen("4_ORDER", 0); SetTag("Selected_URL", 'file:///C:/ASRS_Video/clip125.html')
      on Activate: SetTag("Selected_Medicine", 125)
      on Release: SetTag("ยา 125", 0)
      on Press: SetTag("ยา 125", 1)
   Button "Button_11" at 645,416 size 120x40; TextOff 'Metoprolol'
      on Click: ActivateScreen("4_ORDER", 0); SetTag("Selected_URL", 'file:///C:/ASRS_Video/clip130.html')
      on Activate: SetTag("Selected_Medicine", 130)
      on Release: SetTag("ยา 130", 0)
      on Press: SetTag("ยา 130", 1)
   Button "Button_12" at 24,16 size 94x40; TextOff 'Back'
      on Press: ActivateScreen("2", 0)
   GraphicView "Template_Graphic view_1" at 693,20 size 36x32; Picture "play"
   GraphicView "Template_Graphic view_2" at 27,19 size 36x32; Picture "fast-backward"
   GraphicView "Template_Graphic view_3" at 37,128 size 120x104; Picture "Picture121"
   GraphicView "Template_Graphic view_4" at 191,129 size 120x104; Picture "Picture122"
   GraphicView "Template_Graphic view_5" at 339,129 size 120x104; Picture "Picture123"
   GraphicView "Template_Graphic view_6" at 493,129 size 120x104; Picture "Picture124"
   GraphicView "Template_Graphic view_7" at 645,129 size 120x104; Picture "Picture125"
   GraphicView "Template_Graphic view_8" at 38,305 size 120x104; Picture "Picture126"
   GraphicView "Template_Graphic view_9" at 189,304 size 120x112; Picture "Picture127"
   GraphicView "Template_Graphic view_10" at 351,307 size 96x104; Picture "Picture128"
   GraphicView "Template_Graphic view_11" at 497,304 size 120x112; Picture "Picture129"
   GraphicView "Template_Graphic view_12" at 645,304 size 120x104; Picture "Picture130"
   TextField "Template_Text field_2" at 201,80 size 20x32; Text '3'

screen "4" 800x480, template "Template_2"
   Button "Button_1" at 38,239 size 120x40; TextOff 'Propranolol'
      on Click: ActivateScreen("4_ORDER", 0); SetTag("Selected_URL", 'file:///C:/ASRS_Video/clip131.html')
      on Activate: SetTag("Selected_Medicine", 131)
      on Release: SetTag("ยา 131", 0)
      on Press: SetTag("ยา 131", 1)
   Button "Button_9" at 688,16 size 96x40; TextOff 'Next'
      on Press: ActivateScreen("5", 0)
   Button "Button_10" at 38,415 size 120x40; TextOff 'Aspirin'
      on Click: ActivateScreen("4_ORDER", 0); SetTag("Selected_URL", 'file:///C:/ASRS_Video/clip136.html')
      on Activate: SetTag("Selected_Medicine", 136)
      on Release: SetTag("ยา 136", 0)
      on Press: SetTag("ยา 136", 1)
   Button "Button_2" at 189,240 size 120x40; TextOff 'Carvedilol'
      on Click: ActivateScreen("4_ORDER", 0); SetTag("Selected_URL", 'file:///C:/ASRS_Video/clip132.html')
      on Activate: SetTag("Selected_Medicine", 132)
      on Release: SetTag("ยา 132", 0)
      on Press: SetTag("ยา 132", 1)
   Button "Button_3" at 190,415 size 120x40; TextOff 'Clopidogrel'
      on Click: ActivateScreen("4_ORDER", 0); SetTag("Selected_URL", 'file:///C:/ASRS_Video/clip137.html')
      on Activate: SetTag("Selected_Medicine", 137)
      on Release: SetTag("ยา 137", 0)
      on Press: SetTag("ยา 137", 1)
   Button "Button_4" at 340,240 size 120x40; TextOff 'Digoxin'
      on Click: ActivateScreen("4_ORDER", 0); SetTag("Selected_URL", 'file:///C:/ASRS_Video/clip133.html')
      on Activate: SetTag("Selected_Medicine", 133)
      on Release: SetTag("ยา 133", 0)
      on Press: SetTag("ยา 133", 1)
   Button "Button_5" at 340,416 size 120x40; TextOff 'Warfarin'
      on Click: ActivateScreen("4_ORDER", 0); SetTag("Selected_URL", 'file:///C:/ASRS_Video/clip138.html')
      on Activate: SetTag("Selected_Medicine", 138)
      on Press: SetTag("ยา 138", 1)
   Button "Button_6" at 492,416 size 120x40; TextOff 'Heparin'
      on Click: ActivateScreen("4_ORDER", 0); SetTag("Selected_URL", 'file:///C:/ASRS_Video/clip139.html')
      on Activate: SetTag("Selected_Medicine", 139)
      on Release: SetTag("ยา 139", 0)
      on Press: SetTag("ยา 139", 1)
   Button "Button_7" at 492,240 size 120x40; TextOff 'Isosorbide dinitrate'
      on Click: ActivateScreen("4_ORDER", 0); SetTag("Selected_URL", 'file:///C:/ASRS_Video/clip134.html')
      on Activate: SetTag("Selected_Medicine", 134)
      on Release: SetTag("ยา 134", 0)
      on Press: SetTag("ยา 134", 1)
   Button "Button_8" at 644,240 size 120x40; TextOff 'Nitroglycerin'
      on Click: ActivateScreen("4_ORDER", 0); SetTag("Selected_URL", 'file:///C:/ASRS_Video/clip135.html')
      on Activate: SetTag("Selected_Medicine", 135)
      on Release: SetTag("ยา 135", 0)
      on Press: SetTag("ยา 135", 1)
   Button "Button_11" at 645,416 size 120x40; TextOff 'Enoxaparin'
      on Click: ActivateScreen("4_ORDER", 0); SetTag("Selected_URL", 'file:///C:/ASRS_Video/clip140.html')
      on Activate: SetTag("Selected_Medicine", 140)
      on Release: SetTag("ยา 140", 0)
      on Press: SetTag("ยา 140", 1)
   Button "Button_12" at 24,16 size 94x40; TextOff 'Back'
      on Press: ActivateScreen("3", 0)
   GraphicView "Template_Graphic view_1" at 693,20 size 36x32; Picture "play"
   GraphicView "Template_Graphic view_2" at 27,19 size 36x32; Picture "fast-backward"
   GraphicView "Template_Graphic view_3" at 37,128 size 120x104; Picture "Picture131"
   GraphicView "Template_Graphic view_4" at 191,129 size 120x104; Picture "Picture132"
   GraphicView "Template_Graphic view_5" at 339,129 size 120x104; Picture "Picture133"
   GraphicView "Template_Graphic view_6" at 493,129 size 120x104; Picture "Picture134"
   GraphicView "Template_Graphic view_7" at 645,129 size 120x104; Picture "Picture135"
   GraphicView "Template_Graphic view_8" at 38,305 size 120x104; Picture "Picture136"
   GraphicView "Template_Graphic view_9" at 189,304 size 120x112; Picture "Picture137"
   GraphicView "Template_Graphic view_10" at 351,307 size 96x104; Picture "Picture138"
   GraphicView "Template_Graphic view_11" at 497,304 size 120x112; Picture "Picture139"
   GraphicView "Template_Graphic view_12" at 645,304 size 120x104; Picture "Picture140"
   TextField "Template_Text field_2" at 201,80 size 20x32; Text '4'

screen "5" 800x480, template "Template_2"
   Button "Button_1" at 38,239 size 120x40; TextOff 'Simvastatin'
      on Click: ActivateScreen("4_ORDER", 0); SetTag("Selected_URL", 'file:///C:/ASRS_Video/clip141.html')
      on Activate: SetTag("Selected_Medicine", 141)
      on Release: SetTag("ยา 141", 0)
      on Press: SetTag("ยา 141", 1)
   Button "Button_9" at 688,16 size 96x40; TextOff 'Next'
      on Press: ActivateScreen("6", 0)
   Button "Button_10" at 38,415 size 120x40; TextOff 'Terbutaline'
      on Click: ActivateScreen("4_ORDER", 0); SetTag("Selected_URL", 'file:///C:/ASRS_Video/clip146.html')
      on Activate: SetTag("Selected_Medicine", 146)
      on Release: SetTag("ยา 146", 0)
      on Press: SetTag("ยา 146", 1)
   Button "Button_2" at 189,240 size 120x40; TextOff 'Atorvastatin'
      on Click: ActivateScreen("4_ORDER", 0); SetTag("Selected_URL", 'file:///C:/ASRS_Video/clip142.html')
      on Activate: SetTag("Selected_Medicine", 142)
      on Release: SetTag("ยา 142", 0)
      on Press: SetTag("ยา 142", 1)
   Button "Button_3" at 190,415 size 120x40; TextOff 'Ipratropium bromide'
      on Click: ActivateScreen("4_ORDER", 0); SetTag("Selected_URL", 'file:///C:/ASRS_Video/clip147.html')
      on Activate: SetTag("Selected_Medicine", 147)
      on Release: SetTag("ยา 147", 0)
      on Press: SetTag("ยา 147", 1)
   Button "Button_4" at 340,240 size 120x40; TextOff 'Rosuvastatin'
      on Click: ActivateScreen("4_ORDER", 0); SetTag("Selected_URL", 'file:///C:/ASRS_Video/clip143.html')
      on Activate: SetTag("Selected_Medicine", 143)
      on Release: SetTag("ยา 143", 0)
      on Press: SetTag("ยา 143", 1)
   Button "Button_5" at 340,416 size 120x40; TextOff 'Tiotropium'
      on Click: ActivateScreen("4_ORDER", 0); SetTag("Selected_URL", 'file:///C:/ASRS_Video/clip148.html')
      on Activate: SetTag("Selected_Medicine", 148)
      on Release: SetTag("ยา 148", 0)
      on Press: SetTag("ยา 148", 1)
   Button "Button_6" at 492,416 size 120x40; TextOff 'Budesonide'
      on Click: ActivateScreen("4_ORDER", 0); SetTag("Selected_URL", 'file:///C:/ASRS_Video/clip149.html')
      on Activate: SetTag("Selected_Medicine", 149)
      on Release: SetTag("ยา 149", 0)
      on Press: SetTag("ยา 149", 1)
   Button "Button_7" at 492,240 size 120x40; TextOff 'Gemfibrozil'
      on Click: ActivateScreen("4_ORDER", 0); SetTag("Selected_URL", 'file:///C:/ASRS_Video/clip144.html')
      on Activate: SetTag("Selected_Medicine", 144)
      on Release: SetTag("ยา 144", 0)
      on Press: SetTag("ยา 144", 1)
   Button "Button_8" at 644,240 size 120x40; TextOff 'Salbutamol'
      on Click: ActivateScreen("4_ORDER", 0); SetTag("Selected_URL", 'file:///C:/ASRS_Video/clip145.html')
      on Activate: SetTag("Selected_Medicine", 145)
      on Release: SetTag("ยา 145", 0)
      on Press: SetTag("ยา 145", 1)
   Button "Button_11" at 645,416 size 120x40; TextOff 'Fluticasone'
      on Click: ActivateScreen("4_ORDER", 0); SetTag("Selected_URL", 'file:///C:/ASRS_Video/clip150.html')
      on Activate: SetTag("Selected_Medicine", 150)
      on Release: SetTag("ยา 150", 0)
      on Press: SetTag("ยา 150", 1)
   Button "Button_12" at 24,16 size 94x40; TextOff 'Back'
      on Press: ActivateScreen("4", 0)
   GraphicView "Template_Graphic view_1" at 693,20 size 36x32; Picture "play"
   GraphicView "Template_Graphic view_2" at 27,19 size 36x32; Picture "fast-backward"
   GraphicView "Template_Graphic view_3" at 37,128 size 120x104; Picture "Picture141"
   GraphicView "Template_Graphic view_4" at 191,129 size 120x104; Picture "Picture142"
   GraphicView "Template_Graphic view_5" at 339,129 size 120x104; Picture "Picture143"
   GraphicView "Template_Graphic view_6" at 493,129 size 120x104; Picture "Picture144"
   GraphicView "Template_Graphic view_7" at 645,129 size 120x104; Picture "Picture145"
   GraphicView "Template_Graphic view_8" at 38,305 size 120x104; Picture "Picture146"
   GraphicView "Template_Graphic view_9" at 189,304 size 120x112; Picture "Picture147"
   GraphicView "Template_Graphic view_10" at 351,307 size 96x104; Picture "Picture148"
   GraphicView "Template_Graphic view_11" at 497,304 size 120x112; Picture "Picture149"
   GraphicView "Template_Graphic view_12" at 645,304 size 120x104; Picture "Picture150"
   TextField "Template_Text field_2" at 201,80 size 20x32; Text '5'

screen "6" 800x480, template "Template_2"
   Button "Button_1" at 38,239 size 120x40; TextOff 'Montelukast'
      on Click: ActivateScreen("4_ORDER", 0); SetTag("Selected_URL", 'file:///C:/ASRS_Video/clip151.html')
      on Activate: SetTag("Selected_Medicine", 151)
      on Release: SetTag("ยา 151", 0)
      on Press: SetTag("ยา 151", 1)
   Button "Button_9" at 688,16 size 96x40; TextOff 'Next'
      on Press: ActivateScreen("7", 0)
   Button "Button_10" at 38,415 size 120x40; TextOff 'Dextromethorphan'
      on Click: ActivateScreen("4_ORDER", 0); SetTag("Selected_URL", 'file:///C:/ASRS_Video/clip156.html')
      on Activate: SetTag("Selected_Medicine", 156)
      on Release: SetTag("ยา 156", 0)
      on Press: SetTag("ยา 156", 1)
   Button "Button_2" at 189,240 size 120x40; TextOff 'Theophylline'
      on Click: ActivateScreen("4_ORDER", 0); SetTag("Selected_URL", 'file:///C:/ASRS_Video/clip152.html')
      on Activate: SetTag("Selected_Medicine", 152)
      on Release: SetTag("ยา 152", 0)
      on Press: SetTag("ยา 152", 1)
   Button "Button_3" at 190,415 size 120x40; TextOff 'Chlorpheniramine'
      on Click: ActivateScreen("4_ORDER", 0); SetTag("Selected_URL", 'file:///C:/ASRS_Video/clip157.html')
      on Activate: SetTag("Selected_Medicine", 157)
      on Release: SetTag("ยา 157", 0)
      on Press: SetTag("ยา 157", 1)
   Button "Button_4" at 340,240 size 120x40; TextOff 'Acetylcysteine'
      on Click: ActivateScreen("4_ORDER", 0); SetTag("Selected_URL", 'file:///C:/ASRS_Video/clip153.html')
      on Activate: SetTag("Selected_Medicine", 153)
      on Release: SetTag("ยา 153", 0)
      on Press: SetTag("ยา 153", 1)
   Button "Button_5" at 340,416 size 120x40; TextOff 'Loratadine'
      on Click: ActivateScreen("4_ORDER", 0); SetTag("Selected_URL", 'file:///C:/ASRS_Video/clip158.html')
      on Activate: SetTag("Selected_Medicine", 158)
      on Release: SetTag("ยา 158", 0)
      on Press: SetTag("ยา 158", 1)
   Button "Button_6" at 492,416 size 120x40; TextOff 'Cetirizine'
      on Click: ActivateScreen("4_ORDER", 0); SetTag("Selected_URL", 'file:///C:/ASRS_Video/clip159.html')
      on Activate: SetTag("Selected_Medicine", 159)
      on Release: SetTag("ยา 159", 0)
      on Press: SetTag("ยา 159", 1)
   Button "Button_7" at 492,240 size 120x40; TextOff 'Bromhexine'
      on Click: ActivateScreen("4_ORDER", 0); SetTag("Selected_URL", 'file:///C:/ASRS_Video/clip154.html')
      on Activate: SetTag("Selected_Medicine", 154)
      on Release: SetTag("ยา 154", 0)
      on Press: SetTag("ยา 154", 1)
   Button "Button_8" at 644,240 size 120x40; TextOff 'Ambroxol'
      on Click: ActivateScreen("4_ORDER", 0); SetTag("Selected_URL", 'file:///C:/ASRS_Video/clip155.html')
      on Activate: SetTag("Selected_Medicine", 155)
      on Release: SetTag("ยา 155", 0)
      on Press: SetTag("ยา 155", 1)
   Button "Button_11" at 645,416 size 120x40; TextOff 'Fexofenadine'
      on Click: ActivateScreen("4_ORDER", 0); SetTag("Selected_URL", 'file:///C:/ASRS_Video/clip160.html')
      on Activate: SetTag("Selected_Medicine", 160)
      on Release: SetTag("ยา 160", 0)
      on Press: SetTag("ยา 160", 1)
   Button "Button_12" at 24,16 size 94x40; TextOff 'Back'
      on Press: ActivateScreen("5", 0)
   GraphicView "Template_Graphic view_1" at 693,20 size 36x32; Picture "play"
   GraphicView "Template_Graphic view_2" at 27,19 size 36x32; Picture "fast-backward"
   GraphicView "Template_Graphic view_3" at 37,128 size 120x104; Picture "Picture151"
   GraphicView "Template_Graphic view_4" at 191,129 size 120x104; Picture "Picture152"
   GraphicView "Template_Graphic view_5" at 339,129 size 120x104; Picture "Picture153"
   GraphicView "Template_Graphic view_6" at 493,129 size 120x104; Picture "Picture154"
   GraphicView "Template_Graphic view_7" at 645,129 size 120x104; Picture "Picture155"
   GraphicView "Template_Graphic view_8" at 38,305 size 120x104; Picture "Picture156"
   GraphicView "Template_Graphic view_9" at 189,304 size 120x112; Picture "Picture157"
   GraphicView "Template_Graphic view_10" at 351,307 size 96x104; Picture "Picture158"
   GraphicView "Template_Graphic view_11" at 497,304 size 120x112; Picture "Picture159"
   GraphicView "Template_Graphic view_12" at 645,304 size 120x104; Picture "Picture160"
   TextField "Template_Text field_2" at 201,80 size 20x32; Text '6'

screen "7" 800x480, template "Template_2"
   Button "Button_1" at 38,239 size 120x40; TextOff 'Paracetamol'
      on Click: ActivateScreen("4_ORDER", 0); SetTag("Selected_URL", 'file:///C:/ASRS_Video/clip161.html')
      on Activate: SetTag("Selected_Medicine", 161)
      on Release: SetTag("ยา 161", 0)
      on Press: SetTag("ยา 161", 1)
   Button "Button_9" at 688,16 size 96x40; TextOff 'Next'
      on Press: ActivateScreen("8", 0)
   Button "Button_10" at 38,415 size 120x40; TextOff 'Tramadol'
      on Click: ActivateScreen("4_ORDER", 0); SetTag("Selected_URL", 'file:///C:/ASRS_Video/clip166.html')
      on Activate: SetTag("Selected_Medicine", 166)
      on Release: SetTag("ยา 166", 0)
      on Press: SetTag("ยา 166", 1)
   Button "Button_2" at 189,240 size 120x40; TextOff 'Ibuprofen'
      on Click: ActivateScreen("4_ORDER", 0); SetTag("Selected_URL", 'file:///C:/ASRS_Video/clip162.html')
      on Activate: SetTag("Selected_Medicine", 162)
      on Release: SetTag("ยา 162", 0)
      on Press: SetTag("ยา 162", 1)
   Button "Button_3" at 190,415 size 120x40; TextOff 'Morphine'
      on Click: ActivateScreen("4_ORDER", 0); SetTag("Selected_URL", 'file:///C:/ASRS_Video/clip167.html')
      on Activate: SetTag("Selected_Medicine", 167)
      on Release: SetTag("ยา 167", 0)
      on Press: SetTag("ยา 167", 1)
   Button "Button_4" at 340,240 size 120x40; TextOff 'Diclofenac'
      on Click: ActivateScreen("4_ORDER", 0); SetTag("Selected_URL", 'file:///C:/ASRS_Video/clip163.html')
      on Activate: SetTag("Selected_Medicine", 163)
      on Release: SetTag("ยา 163", 0)
      on Press: SetTag("ยา 163", 1)
   Button "Button_5" at 340,416 size 120x40; TextOff 'Codeine'
      on Click: ActivateScreen("4_ORDER", 0); SetTag("Selected_URL", 'file:///C:/ASRS_Video/clip168.html')
      on Activate: SetTag("Selected_Medicine", 168)
      on Release: SetTag("ยา 168", 0)
      on Press: SetTag("ยา 168", 1)
   Button "Button_6" at 492,416 size 120x40; TextOff 'Gabapentin'
      on Click: ActivateScreen("4_ORDER", 0); SetTag("Selected_URL", 'file:///C:/ASRS_Video/clip169.html')
      on Activate: SetTag("Selected_Medicine", 169)
      on Release: SetTag("ยา 169", 0)
      on Press: SetTag("ยา 169", 1)
   Button "Button_7" at 492,240 size 120x40; TextOff 'Naproxen'
      on Click: ActivateScreen("4_ORDER", 0); SetTag("Selected_URL", 'file:///C:/ASRS_Video/clip164.html')
      on Activate: SetTag("Selected_Medicine", 164)
      on Release: SetTag("ยา 164", 0)
      on Press: SetTag("ยา 164", 1)
   Button "Button_8" at 644,240 size 120x40; TextOff 'Celecoxib'
      on Click: ActivateScreen("4_ORDER", 0); SetTag("Selected_URL", 'file:///C:/ASRS_Video/clip165.html')
      on Activate: SetTag("Selected_Medicine", 165)
      on Release: SetTag("ยา 165", 0)
      on Press: SetTag("ยา 165", 1)
   Button "Button_11" at 645,416 size 120x40; TextOff 'Pregabalin'
      on Click: ActivateScreen("4_ORDER", 0); SetTag("Selected_URL", 'file:///C:/ASRS_Video/clip170.html')
      on Activate: SetTag("Selected_Medicine", 170)
      on Release: SetTag("ยา 170", 0)
      on Press: SetTag("ยา 170", 1)
   Button "Button_12" at 24,16 size 94x40; TextOff 'Back'
      on Press: ActivateScreen("6", 0)
   GraphicView "Template_Graphic view_1" at 693,20 size 36x32; Picture "play"
   GraphicView "Template_Graphic view_2" at 27,19 size 36x32; Picture "fast-backward"
   GraphicView "Template_Graphic view_3" at 37,128 size 120x104; Picture "Picture161"
   GraphicView "Template_Graphic view_4" at 191,129 size 120x104; Picture "Picture162"
   GraphicView "Template_Graphic view_5" at 339,129 size 120x104; Picture "Picture163"
   GraphicView "Template_Graphic view_6" at 493,129 size 120x104; Picture "Picture164"
   GraphicView "Template_Graphic view_7" at 645,129 size 120x104; Picture "Picture165"
   GraphicView "Template_Graphic view_8" at 38,305 size 120x104; Picture "Picture166"
   GraphicView "Template_Graphic view_9" at 189,304 size 120x112; Picture "Picture167"
   GraphicView "Template_Graphic view_10" at 351,307 size 96x104; Picture "Picture168"
   GraphicView "Template_Graphic view_11" at 497,304 size 120x112; Picture "Picture169"
   GraphicView "Template_Graphic view_12" at 645,304 size 120x104; Picture "Picture170"
   TextField "Template_Text field_2" at 201,80 size 20x32; Text '7'

screen "8" 800x480, template "Template_2"
   Button "Button_1" at 38,239 size 120x40; TextOff 'Amitriptyline'
      on Click: ActivateScreen("4_ORDER", 0); SetTag("Selected_URL", 'file:///C:/ASRS_Video/clip171.html')
      on Activate: SetTag("Selected_Medicine", 171)
      on Release: SetTag("ยา 171", 0)
      on Press: SetTag("ยา 171", 1)
   Button "Button_10" at 38,415 size 120x40; TextOff 'Lorazepam'
      on Click: ActivateScreen("4_ORDER", 0); SetTag("Selected_URL", 'file:///C:/ASRS_Video/clip176.html')
      on Activate: SetTag("Selected_Medicine", 176)
      on Release: SetTag("ยา 176", 0)
      on Press: SetTag("ยา 176", 1)
   Button "Button_2" at 189,240 size 120x40; TextOff 'Nortriptyline'
      on Click: ActivateScreen("4_ORDER", 0); SetTag("Selected_URL", 'file:///C:/ASRS_Video/clip172.html')
      on Activate: SetTag("Selected_Medicine", 172)
      on Release: SetTag("ยา 172", 0)
      on Press: SetTag("ยา 172", 1)
   Button "Button_3" at 190,415 size 120x40; TextOff 'Alprazolam'
      on Click: ActivateScreen("4_ORDER", 0); SetTag("Selected_URL", 'file:///C:/ASRS_Video/clip177.html')
      on Activate: SetTag("Selected_Medicine", 177)
      on Release: SetTag("ยา 177", 0)
      on Press: SetTag("ยา 177", 1)
   Button "Button_4" at 340,240 size 120x40; TextOff 'Fluoxetine'
      on Click: ActivateScreen("4_ORDER", 0); SetTag("Selected_URL", 'file:///C:/ASRS_Video/clip173.html')
      on Activate: SetTag("Selected_Medicine", 173)
      on Release: SetTag("ยา 173", 0)
      on Press: SetTag("ยา 173", 1)
   Button "Button_5" at 340,416 size 120x40; TextOff 'Clonazepam'
      on Click: ActivateScreen("4_ORDER", 0); SetTag("Selected_URL", 'file:///C:/ASRS_Video/clip178.html')
      on Activate: SetTag("Selected_Medicine", 178)
      on Release: SetTag("ยา 178", 0)
      on Press: SetTag("ยา 178", 1)
   Button "Button_6" at 492,416 size 120x40; TextOff 'Phenytoin'
      on Click: ActivateScreen("4_ORDER", 0); SetTag("Selected_URL", 'file:///C:/ASRS_Video/clip179.html')
      on Activate: SetTag("Selected_Medicine", 179)
      on Release: SetTag("ยา 179", 0)
      on Press: SetTag("ยา 179", 1)
   Button "Button_7" at 492,240 size 120x40; TextOff 'Sertraline'
      on Click: ActivateScreen("4_ORDER", 0); SetTag("Selected_URL", 'file:///C:/ASRS_Video/clip174.html')
      on Activate: SetTag("Selected_Medicine", 174)
      on Release: SetTag("ยา 174", 0)
      on Press: SetTag("ยา 174", 1)
   Button "Button_8" at 644,240 size 120x40; TextOff 'Diazepam'
      on Click: ActivateScreen("4_ORDER", 0); SetTag("Selected_URL", 'file:///C:/ASRS_Video/clip175.html')
      on Activate: SetTag("Selected_Medicine", 175)
      on Release: SetTag("ยา 175", 0)
      on Press: SetTag("ยา 175", 1)
   Button "Button_11" at 645,416 size 120x40; TextOff 'Sodium valproate'
      on Click: ActivateScreen("4_ORDER", 0); SetTag("Selected_URL", 'file:///C:/ASRS_Video/clip180.html')
      on Activate: SetTag("Selected_Medicine", 180)
      on Release: SetTag("ยา 180", 0)
      on Press: SetTag("ยา 180", 1)
   Button "Button_12" at 24,16 size 94x40; TextOff 'Back'
      on Press: ActivateScreen("7", 0)
   Button "Button_9" at 688,16 size 96x40; TextOff 'Next'
      on Press: ActivateScreen("9", 0)
   GraphicView "Template_Graphic view_2" at 27,19 size 36x32; Picture "fast-backward"
   GraphicView "Template_Graphic view_1" at 693,20 size 36x32; Picture "play"
   GraphicView "Template_Graphic view_3" at 37,128 size 120x104; Picture "Picture171"
   GraphicView "Template_Graphic view_4" at 191,129 size 120x104; Picture "Picture172"
   GraphicView "Template_Graphic view_5" at 339,129 size 120x104; Picture "Picture173"
   GraphicView "Template_Graphic view_6" at 493,129 size 120x104; Picture "Picture174"
   GraphicView "Template_Graphic view_7" at 645,129 size 120x104; Picture "Picture175"
   GraphicView "Template_Graphic view_8" at 38,305 size 120x104; Picture "Picture176"
   GraphicView "Template_Graphic view_9" at 189,304 size 120x112; Picture "Picture177"
   GraphicView "Template_Graphic view_10" at 351,307 size 96x104; Picture "Picture178"
   GraphicView "Template_Graphic view_11" at 497,304 size 120x112; Picture "Picture179"
   GraphicView "Template_Graphic view_12" at 645,304 size 120x104; Picture "Picture180"
   TextField "Template_Text field_2" at 201,80 size 20x32; Text '8'

